   // ---------- 网络 17 ----------
   // 标题：请开始换夹具...
   // 含义：将 (#ChangeTool.S15 AND #StatusIn.do_ChgGrp_Pos) OR (#ChangeTool.S15 AND #ChangeTool.S17) 赋给 #ChangeTool.S17
   #ChangeTool.S17 := (#ChangeTool.S15 AND #StatusIn.do_ChgGrp_Pos) OR (#ChangeTool.S15 AND #ChangeTool.S17);
   // 含义：将 #ChangeTool.S15 AND NOT (#ChangeTool.S17) 赋给 "DB1146_PromptFree".Public.do_ChgGrp_Pos
   "DB1146_PromptFree".Public.do_ChgGrp_Pos := #ChangeTool.S15 AND NOT (#ChangeTool.S17);

   // ---------- 网络 18 ----------
   // 标题：快换盘锁紧 254放爪 253取爪
   // 含义：条件 ((#ChangeTool.S17 AND NOT (#ChangeTool.S19)) AND ("DB1080_Component".Robot.CTRL_IN.ProgNo = 253)) 成立时，将 TRUE 传送到 "DB1081_ValveCall".ST01.Z07.ExtAuto
   IF ((#ChangeTool.S17 AND NOT (#ChangeTool.S19)) AND ("DB1080_Component".Robot.CTRL_IN.ProgNo = 253)) THEN
       "DB1081_ValveCall".ST01.Z07.ExtAuto := TRUE;
   END_IF;
   // 含义：条件 ((#ChangeTool.S17 AND NOT (#ChangeTool.S19)) AND ("DB1080_Component".Robot.CTRL_IN.ProgNo = 254)) 成立时，将 TRUE 传送到 "DB1081_ValveCall".ST01.Z07.RetAuto
   IF ((#ChangeTool.S17 AND NOT (#ChangeTool.S19)) AND ("DB1080_Component".Robot.CTRL_IN.ProgNo = 254)) THEN
       "DB1081_ValveCall".ST01.Z07.RetAuto := TRUE;
   END_IF;
   // 含义：条件 #ChangeTool.S17 AND NOT (#ChangeTool.S19) 成立时，将 TRUE 传送到 "DB1060_AutoStep".Status.FirstStart
   IF #ChangeTool.S17 AND NOT (#ChangeTool.S19) THEN
       "DB1060_AutoStep".Status.FirstStart := TRUE;
   END_IF;
   // 含义：将 (((#ChangeTool.S17 AND ("DB1080_Component".Robot.CTRL_IN.ProgNo = 253))) AND "DB1081_ValveCall".ST01.Z07.ExtPos) OR (((#ChangeTool.S17 AND ("DB1080_Component".Robot.CTRL_IN.ProgNo = 254))) AND "DB1081_ValveCall".ST01.Z07.RetPos) OR (#ChangeTool.S17 AND #ChangeTool.S19) 赋给 #ChangeTool.S19
   #ChangeTool.S19 := (((#ChangeTool.S17 AND ("DB1080_Component".Robot.CTRL_IN.ProgNo = 253))) AND "DB1081_ValveCall".ST01.Z07.ExtPos) OR (((#ChangeTool.S17 AND ("DB1080_Component".Robot.CTRL_IN.ProgNo = 254))) AND "DB1081_ValveCall".ST01.Z07.RetPos) OR (#ChangeTool.S17 AND #ChangeTool.S19);

   // ---------- 网络 19 ----------
   // 标题：换爪完成确认
   // 含义：将 #ChangeTool.S19 AND NOT (#ChangeTool.S20) 赋给 #CmdOut.di_ChgGrp_Ack
   #CmdOut.di_ChgGrp_Ack := #ChangeTool.S19 AND NOT (#ChangeTool.S20);
   // 含义：将 #ChangeTool.S19 AND NOT (#ChangeTool.S20) 赋给 "DB1146_PromptFree".Public.do_ChgGrp_Act
   "DB1146_PromptFree".Public.do_ChgGrp_Act := #ChangeTool.S19 AND NOT (#ChangeTool.S20);
   // 含义：条件 (#ChangeTool.S19 AND NOT (#ChangeTool.S20)) AND NOT ("IToolAtPos") 成立时，将 TRUE 传送到 "DB1081_ValveCall".ST01.Z07.VentValveAuto
   IF (#ChangeTool.S19 AND NOT (#ChangeTool.S20)) AND NOT ("IToolAtPos") THEN
       "DB1081_ValveCall".ST01.Z07.VentValveAuto := TRUE;
   END_IF;
   // 含义：条件 #ChangeTool.S19 AND NOT (#ChangeTool.S20) 成立时，将 TRUE 传送到 "DB1081_ValveCall".ST01.Z08.RetAuto
   IF #ChangeTool.S19 AND NOT (#ChangeTool.S20) THEN
       "DB1081_ValveCall".ST01.Z08.RetAuto := TRUE;
   END_IF;
   // 含义：将 (#ChangeTool.S19 AND #StatusIn.do_ChgGrp_Don) OR (#ChangeTool.S19 AND #ChangeTool.S20) 赋给 #ChangeTool.S20
   #ChangeTool.S20 := (#ChangeTool.S19 AND #StatusIn.do_ChgGrp_Don) OR (#ChangeTool.S19 AND #ChangeTool.S20);

   // ---------- 网络 20 ----------
   // 标题：夹具库枪位置不正确！
   // 注释：M29.0常1临时屏蔽I6.0信号 20230911
   // 含义：将 (((((#ChangeTool.S20 AND ("DB1080_Component".Robot.CTRL_IN.ProgNo = 254))) AND (#CmdOut.gi_ToolPosNo = 1))) AND NOT (#Aux.AStation_ToolAtPosT.Q)) OR (((((#ChangeTool.S20 AND ("DB1080_Component".Robot.CTRL_IN.ProgNo = 254))) AND (#CmdOut.gi_ToolPosNo = 2))) AND NOT (#Aux.BStation_ToolAtPosT.Q)) 赋给 "DB1148_PromptBeeper".ST01.PutToolPosNotOk
   "DB1148_PromptBeeper".ST01.PutToolPosNotOk := (((((#ChangeTool.S20 AND ("DB1080_Component".Robot.CTRL_IN.ProgNo = 254))) AND (#CmdOut.gi_ToolPosNo = 1))) AND NOT (#Aux.AStation_ToolAtPosT.Q)) OR (((((#ChangeTool.S20 AND ("DB1080_Component".Robot.CTRL_IN.ProgNo = 254))) AND (#CmdOut.gi_ToolPosNo = 2))) AND NOT (#Aux.BStation_ToolAtPosT.Q));
   // 含义：将 (((((#ChangeTool.S20 AND ("DB1080_Component".Robot.CTRL_IN.ProgNo = 254))) AND (#CmdOut.gi_ToolPosNo = 1))) AND #Aux.AStation_ToolAtPosT.Q) OR (((((#ChangeTool.S20 AND ("DB1080_Component".Robot.CTRL_IN.ProgNo = 254))) AND (#CmdOut.gi_ToolPosNo = 2))) AND #Aux.BStation_ToolAtPosT.Q) OR ((((#ChangeTool.S20 AND ("DB1080_Component".Robot.CTRL_IN.ProgNo = 253))) AND "DB1081_ValveCall".ST01.Z07.ExtPos) AND "IToolAtPos") OR (#ChangeTool.S20 AND #ChangeTool.S22) 赋给 #ChangeTool.S22
   #ChangeTool.S22 := (((((#ChangeTool.S20 AND ("DB1080_Component".Robot.CTRL_IN.ProgNo = 254))) AND (#CmdOut.gi_ToolPosNo = 1))) AND #Aux.AStation_ToolAtPosT.Q) OR (((((#ChangeTool.S20 AND ("DB1080_Component".Robot.CTRL_IN.ProgNo = 254))) AND (#CmdOut.gi_ToolPosNo = 2))) AND #Aux.BStation_ToolAtPosT.Q) OR ((((#ChangeTool.S20 AND ("DB1080_Component".Robot.CTRL_IN.ProgNo = 253))) AND "DB1081_ValveCall".ST01.Z07.ExtPos) AND "IToolAtPos") OR (#ChangeTool.S20 AND #ChangeTool.S22);

   // ---------- 网络 21 ----------
   // 标题：防尘盖夹紧缸
   // 含义：条件 ((((#ChangeTool.S22 AND NOT (#ChangeTool.S23)) AND ("DB1080_Component".Robot.CTRL_IN.ProgNo <> 254))) OR ((#ChangeTool.S22 AND NOT (#ChangeTool.S23)) AND TRUE)) AND #Aux.AStation_ToolAtPosT.Q 成立时，将 TRUE 传送到 "DB1081_ValveCall".ST01.Z03.RetAuto
   IF ((((#ChangeTool.S22 AND NOT (#ChangeTool.S23)) AND ("DB1080_Component".Robot.CTRL_IN.ProgNo <> 254))) OR ((#ChangeTool.S22 AND NOT (#ChangeTool.S23)) AND TRUE)) AND #Aux.AStation_ToolAtPosT.Q THEN
       "DB1081_ValveCall".ST01.Z03.RetAuto := TRUE;
   END_IF;
   // 含义：条件 ((((#ChangeTool.S22 AND NOT (#ChangeTool.S23)) AND ("DB1080_Component".Robot.CTRL_IN.ProgNo <> 254))) OR ((#ChangeTool.S22 AND NOT (#ChangeTool.S23)) AND TRUE)) AND #Aux.BStation_ToolAtPosT.Q 成立时，将 TRUE 传送到 "DB1081_ValveCall".ST01.Z04.RetAuto
   IF ((((#ChangeTool.S22 AND NOT (#ChangeTool.S23)) AND ("DB1080_Component".Robot.CTRL_IN.ProgNo <> 254))) OR ((#ChangeTool.S22 AND NOT (#ChangeTool.S23)) AND TRUE)) AND #Aux.BStation_ToolAtPosT.Q THEN
       "DB1081_ValveCall".ST01.Z04.RetAuto := TRUE;
   END_IF;
   // 含义：将 (((#ChangeTool.S22 AND "DB1081_ValveCall".ST01.Z03.RetPos) OR (#ChangeTool.S22 AND NOT (#Aux.AStation_ToolAtPosT.Q))) AND "DB1081_ValveCall".ST01.Z04.RetPos) OR (((#ChangeTool.S22 AND "DB1081_ValveCall".ST01.Z03.RetPos) OR (#ChangeTool.S22 AND NOT (#Aux.AStation_ToolAtPosT.Q))) AND NOT (#Aux.BStation_ToolAtPosT.Q)) OR ((#ChangeTool.S22 AND ("DB1080_Component".Robot.CTRL_IN.ProgNo = 254))) OR (#ChangeTool.S22 AND #ChangeTool.S23) 赋给 #ChangeTool.S23
   #ChangeTool.S23 := (((#ChangeTool.S22 AND "DB1081_ValveCall".ST01.Z03.RetPos) OR (#ChangeTool.S22 AND NOT (#Aux.AStation_ToolAtPosT.Q))) AND "DB1081_ValveCall".ST01.Z04.RetPos) OR (((#ChangeTool.S22 AND "DB1081_ValveCall".ST01.Z03.RetPos) OR (#ChangeTool.S22 AND NOT (#Aux.AStation_ToolAtPosT.Q))) AND NOT (#Aux.BStation_ToolAtPosT.Q)) OR ((#ChangeTool.S22 AND ("DB1080_Component".Robot.CTRL_IN.ProgNo = 254))) OR (#ChangeTool.S22 AND #ChangeTool.S23);

   // ---------- 网络 22 ----------
   // 标题：TaskDone
   // 含义：条件 ((#ChangeTool.S23 OR #ChangeTool.ErrEnd OR #ChangeTool.ByPass) AND NOT (#ChangeTool.S25)) AND NOT (#ChangeTool.ErrEnd) 成立时，将 TRUE 传送到 #ChangeTool.TaskIO
   IF ((#ChangeTool.S23 OR #ChangeTool.ErrEnd OR #ChangeTool.ByPass) AND NOT (#ChangeTool.S25)) AND NOT (#ChangeTool.ErrEnd) THEN
       #ChangeTool.TaskIO := TRUE;
   END_IF;
   // 含义：条件 ((#ChangeTool.S23 OR #ChangeTool.ErrEnd OR #ChangeTool.ByPass) AND NOT (#ChangeTool.S25)) AND #ChangeTool.ErrEnd 成立时，将 TRUE 传送到 #ChangeTool.TaskNIO
   IF ((#ChangeTool.S23 OR #ChangeTool.ErrEnd OR #ChangeTool.ByPass) AND NOT (#ChangeTool.S25)) AND #ChangeTool.ErrEnd THEN
       #ChangeTool.TaskNIO := TRUE;
   END_IF;
   // 含义：将 #ChangeTool.S23 OR #ChangeTool.ErrEnd OR #ChangeTool.ByPass 赋给 #ChangeTool.S25
   #ChangeTool.S25 := #ChangeTool.S23 OR #ChangeTool.ErrEnd OR #ChangeTool.ByPass;

   // ---------- 网络 23 ----------
   // 标题：结束
   // 含义：将 (#ChangeTool.S25 OR #ChangeTool.ErrEnd) AND NOT (#ChangeTool.StartCmd) 赋给 #ChangeTool.StepEnd
   #ChangeTool.StepEnd := (#ChangeTool.S25 OR #ChangeTool.ErrEnd) AND NOT (#ChangeTool.StartCmd);
   // 含义：将 #ChangeTool.S25 OR #ChangeTool.ErrEnd 赋给 #ChangeTool.TaskDone
   #ChangeTool.TaskDone := #ChangeTool.S25 OR #ChangeTool.ErrEnd;

   // ---------- 网络 24 ----------
   // 含义：将 FALSE 赋给 #ChangeTool.StartCmd
   #ChangeTool.StartCmd := FALSE;

   // ---------- 网络 25 ----------
   // （空白网络）

   // ---------- 网络 26 ----------
   // 标题：本工位必须要做(可能条件暂时不满足)
   // 含义：将 (((((#Ctrl_Out.RobotAction = 0) AND #Aux.ToolAtPos) AND "ManMode_M") AND ("DB1900_Communication_PC".Recv.ChooseProgNo = 4))) OR (((((#Ctrl_Out.RobotAction = 0) AND #Aux.ToolAtPos) AND "ManMode_M") AND ("DB1900_Communication_PC".Recv.ChooseProgNo = 5))) OR (((#Ctrl_Out.RobotAction = 0) AND #Aux.ToolAtPos) AND "ASMMode_M") 赋给 #CheckBit.OKToStart
   #CheckBit.OKToStart := (((((#Ctrl_Out.RobotAction = 0) AND #Aux.ToolAtPos) AND "ManMode_M") AND ("DB1900_Communication_PC".Recv.ChooseProgNo = 4))) OR (((((#Ctrl_Out.RobotAction = 0) AND #Aux.ToolAtPos) AND "ManMode_M") AND ("DB1900_Communication_PC".Recv.ChooseProgNo = 5))) OR (((#Ctrl_Out.RobotAction = 0) AND #Aux.ToolAtPos) AND "ASMMode_M");
   // 含义：条件 "DB1900_Communication_PC".Recv.CheckAiguilleTPPB AND "ManMode_M" 成立时，将 TRUE 传送到 #CheckBit.StartCmd
   IF "DB1900_Communication_PC".Recv.CheckAiguilleTPPB AND "ManMode_M" THEN
       #CheckBit.StartCmd := TRUE;
   END_IF;

   // ---------- 网络 27 ----------
   // 标题：*********************************检查批头Start*************************************
   // 含义：将 (((((((#CheckBit.StartCmd AND #CheckBit.OKToStart) OR #CheckBit.StepStart) AND "AllMode_M") AND "DB1900_Communication_PC".Recv.Z05RetTPPB) AND ("DB1900_Communication_PC".Recv.Current_2 < 0.5))) AND NOT ("DB1040_HomePos".Status.Running)) AND NOT (#CheckBit.StepEnd) 赋给 #CheckBit.StepStart
   #CheckBit.StepStart := (((((((#CheckBit.StartCmd AND #CheckBit.OKToStart) OR #CheckBit.StepStart) AND "AllMode_M") AND "DB1900_Communication_PC".Recv.Z05RetTPPB) AND ("DB1900_Communication_PC".Recv.Current_2 < 0.5))) AND NOT ("DB1040_HomePos".Status.Running)) AND NOT (#CheckBit.StepEnd);
   // 含义：将 (((((((#CheckBit.StartCmd AND #CheckBit.OKToStart) OR #CheckBit.StepStart) AND "AllMode_M") AND "DB1900_Communication_PC".Recv.Z05RetTPPB) AND ("DB1900_Communication_PC".Recv.Current_2 < 0.5))) AND NOT ("DB1040_HomePos".Status.Running)) AND NOT (#CheckBit.StepEnd) 赋给 #CheckBit.Busy
   #CheckBit.Busy := (((((((#CheckBit.StartCmd AND #CheckBit.OKToStart) OR #CheckBit.StepStart) AND "AllMode_M") AND "DB1900_Communication_PC".Recv.Z05RetTPPB) AND ("DB1900_Communication_PC".Recv.Current_2 < 0.5))) AND NOT ("DB1040_HomePos".Status.Running)) AND NOT (#CheckBit.StepEnd);
   // 含义：将 (((((((#CheckBit.StartCmd AND #CheckBit.OKToStart) OR #CheckBit.StepStart) AND "AllMode_M") AND "DB1900_Communication_PC".Recv.Z05RetTPPB) AND ("DB1900_Communication_PC".Recv.Current_2 < 0.5))) AND NOT ("DB1040_HomePos".Status.Running)) AND NOT (#CheckBit.StepEnd) 赋给 "DB1900_Communication_PC".Send.RobotCheck
   "DB1900_Communication_PC".Send.RobotCheck := (((((((#CheckBit.StartCmd AND #CheckBit.OKToStart) OR #CheckBit.StepStart) AND "AllMode_M") AND "DB1900_Communication_PC".Recv.Z05RetTPPB) AND ("DB1900_Communication_PC".Recv.Current_2 < 0.5))) AND NOT ("DB1040_HomePos".Status.Running)) AND NOT (#CheckBit.StepEnd);
   // 含义：条件 NOT ((((((((#CheckBit.StartCmd AND #CheckBit.OKToStart) OR #CheckBit.StepStart) AND "AllMode_M") AND "DB1900_Communication_PC".Recv.Z05RetTPPB) AND ("DB1900_Communication_PC".Recv.Current_2 < 0.5))) AND NOT ("DB1040_HomePos".Status.Running)) AND NOT (#CheckBit.StepEnd)) 成立时，将 FALSE 传送到 #CheckBit.ErrEnd
   IF NOT ((((((((#CheckBit.StartCmd AND #CheckBit.OKToStart) OR #CheckBit.StepStart) AND "AllMode_M") AND "DB1900_Communication_PC".Recv.Z05RetTPPB) AND ("DB1900_Communication_PC".Recv.Current_2 < 0.5))) AND NOT ("DB1040_HomePos".Status.Running)) AND NOT (#CheckBit.StepEnd)) THEN
       #CheckBit.ErrEnd := FALSE;
   END_IF;
   // 含义：条件 NOT ((((((((#CheckBit.StartCmd AND #CheckBit.OKToStart) OR #CheckBit.StepStart) AND "AllMode_M") AND "DB1900_Communication_PC".Recv.Z05RetTPPB) AND ("DB1900_Communication_PC".Recv.Current_2 < 0.5))) AND NOT ("DB1040_HomePos".Status.Running)) AND NOT (#CheckBit.StepEnd)) 成立时，将 FALSE 传送到 "DB1148_PromptBeeper".Public.ScrLenFault
   IF NOT ((((((((#CheckBit.StartCmd AND #CheckBit.OKToStart) OR #CheckBit.StepStart) AND "AllMode_M") AND "DB1900_Communication_PC".Recv.Z05RetTPPB) AND ("DB1900_Communication_PC".Recv.Current_2 < 0.5))) AND NOT ("DB1040_HomePos".Status.Running)) AND NOT (#CheckBit.StepEnd)) THEN
       "DB1148_PromptBeeper".Public.ScrLenFault := FALSE;
   END_IF;
   // 含义：条件 NOT ((((((((#CheckBit.StartCmd AND #CheckBit.OKToStart) OR #CheckBit.StepStart) AND "AllMode_M") AND "DB1900_Communication_PC".Recv.Z05RetTPPB) AND ("DB1900_Communication_PC".Recv.Current_2 < 0.5))) AND NOT ("DB1040_HomePos".Status.Running)) AND NOT (#CheckBit.StepEnd)) 成立时，将 FALSE 传送到 #CmdOut.di_ChkScrew_Ack
   IF NOT ((((((((#CheckBit.StartCmd AND #CheckBit.OKToStart) OR #CheckBit.StepStart) AND "AllMode_M") AND "DB1900_Communication_PC".Recv.Z05RetTPPB) AND ("DB1900_Communication_PC".Recv.Current_2 < 0.5))) AND NOT ("DB1040_HomePos".Status.Running)) AND NOT (#CheckBit.StepEnd)) THEN
       #CmdOut.di_ChkScrew_Ack := FALSE;
   END_IF;

   // ---------- 网络 28 ----------
   // 标题：初始化
   // 含义：条件 (#CheckBit.StepStart AND NOT (#CheckBit.ErrEnd)) AND NOT (#CheckBit.S1) 成立时，将 FALSE 传送到 #CheckBit.TaskIO
   IF (#CheckBit.StepStart AND NOT (#CheckBit.ErrEnd)) AND NOT (#CheckBit.S1) THEN
       #CheckBit.TaskIO := FALSE;
   END_IF;
   // 含义：条件 (#CheckBit.StepStart AND NOT (#CheckBit.ErrEnd)) AND NOT (#CheckBit.S1) 成立时，将 FALSE 传送到 #CheckBit.TaskNIO
   IF (#CheckBit.StepStart AND NOT (#CheckBit.ErrEnd)) AND NOT (#CheckBit.S1) THEN
       #CheckBit.TaskNIO := FALSE;
   END_IF;
   // 含义：将 #CheckBit.StepStart AND NOT (#CheckBit.ErrEnd) 赋给 #CheckBit.S1
   #CheckBit.S1 := #CheckBit.StepStart AND NOT (#CheckBit.ErrEnd);

   // ---------- 网络 29 ----------
   // 标题：判断条件
   // 含义：当 #CheckBit.S1 为 TRUE 时置位 #CheckBit.S2，否则复位（触点→线圈）
   IF #CheckBit.S1 THEN
       #CheckBit.S2 := TRUE;
   ELSE
       #CheckBit.S2 := FALSE;
   END_IF;

   // ---------- 网络 30 ----------
   // 标题：电源夹具ID号错误，请检查夹具！
   // 含义：将 (#CheckBit.S2 AND #Aux.ToolAtPos) OR (#CheckBit.S2 AND #CheckBit.S5) 赋给 #CheckBit.S5
   #CheckBit.S5 := (#CheckBit.S2 AND #Aux.ToolAtPos) OR (#CheckBit.S2 AND #CheckBit.S5);

   // ---------- 网络 31 ----------
   // 标题：推力气缸
   // 含义：条件 #CheckBit.S5 AND NOT (#CheckBit.S7) 成立时，将 TRUE 传送到 "DB1081_ValveCall".ST01.Z01.ExtAuto
   IF #CheckBit.S5 AND NOT (#CheckBit.S7) THEN
       "DB1081_ValveCall".ST01.Z01.ExtAuto := TRUE;
   END_IF;
   // 含义：条件 #CheckBit.S5 AND NOT (#CheckBit.S7) 成立时，将 TRUE 传送到 "DB1081_ValveCall".ST01.Z02.VentValveAuto
   IF #CheckBit.S5 AND NOT (#CheckBit.S7) THEN
       "DB1081_ValveCall".ST01.Z02.VentValveAuto := TRUE;
   END_IF;
   // 含义：条件 #CheckBit.S5 AND NOT (#CheckBit.S7) 成立时，将 TRUE 传送到 "DB1081_ValveCall".ST01.Z05.RetAuto
   IF #CheckBit.S5 AND NOT (#CheckBit.S7) THEN
       "DB1081_ValveCall".ST01.Z05.RetAuto := TRUE;
   END_IF;
   // 含义：条件 #CheckBit.S5 AND NOT (#CheckBit.S7) 成立时，将 TRUE 传送到 "DB1081_ValveCall".ST01.Z06.RetAuto
   IF #CheckBit.S5 AND NOT (#CheckBit.S7) THEN
       "DB1081_ValveCall".ST01.Z06.RetAuto := TRUE;
   END_IF;
   // 含义：条件 (((#CheckBit.S5 AND NOT (#CheckBit.S7)) AND (#CmdOut.gi_ToolTypeNo = 13))) AND TRUE 成立时，将 FALSE 传送到 "QCamCoverExt"
   IF (((#CheckBit.S5 AND NOT (#CheckBit.S7)) AND (#CmdOut.gi_ToolTypeNo = 13))) AND TRUE THEN
       "QCamCoverExt" := FALSE;
   END_IF;
   // 含义：条件 (((#CheckBit.S5 AND NOT (#CheckBit.S7)) AND (#CmdOut.gi_ToolTypeNo = 13))) AND TRUE 成立时，将 TRUE 传送到 "QCamCoverRet"
   IF (((#CheckBit.S5 AND NOT (#CheckBit.S7)) AND (#CmdOut.gi_ToolTypeNo = 13))) AND TRUE THEN
       "QCamCoverRet" := TRUE;
   END_IF;
   // 含义：条件 #CheckBit.S5 AND NOT (#CheckBit.S7) 成立时，将 TRUE 传送到 "DB1081_ValveCall".ST01.Z08.ExtAuto
   IF #CheckBit.S5 AND NOT (#CheckBit.S7) THEN
       "DB1081_ValveCall".ST01.Z08.ExtAuto := TRUE;
   END_IF;
   // 含义：条件 #CheckBit.S5 AND NOT (#CheckBit.S7) 成立时，将 0.15 传送到 "DB1080_Component".Aux.Pressure
   IF #CheckBit.S5 AND NOT (#CheckBit.S7) THEN
       "DB1080_Component".Aux.Pressure := 0.15;
   END_IF;
   // 含义：将 ((((#CheckBit.S5 AND "DB1900_Communication_PC".Recv.ParaWriteDone) AND "DB1081_ValveCall".ST01.Z05.RetPos) AND "DB1081_ValveCall".ST01.Z06.RetPos) AND "IZ02ExtPos") OR (#CheckBit.S5 AND #CheckBit.S7) 赋给 #CheckBit.S7
   #CheckBit.S7 := ((((#CheckBit.S5 AND "DB1900_Communication_PC".Recv.ParaWriteDone) AND "DB1081_ValveCall".ST01.Z05.RetPos) AND "DB1081_ValveCall".ST01.Z06.RetPos) AND "IZ02ExtPos") OR (#CheckBit.S5 AND #CheckBit.S7);

   // ---------- 网络 32 ----------
   // 标题：数据写入 零点推力压缩量传递
   // 含义：条件 #CheckBit.S7 AND NOT (#CheckBit.S9) 成立时，将 "DB1900_Communication_PC".Para.ZeroPos 传送到 #Aux.ZeroPos
   IF #CheckBit.S7 AND NOT (#CheckBit.S9) THEN
       #Aux.ZeroPos := "DB1900_Communication_PC".Para.ZeroPos;
   END_IF;
   // 含义：当 #CheckBit.S7 为 TRUE 时置位 #CheckBit.S9，否则复位（触点→线圈）
   IF #CheckBit.S7 THEN
       #CheckBit.S9 := TRUE;
   ELSE
       #CheckBit.S9 := FALSE;
   END_IF;

   // ---------- 网络 33 ----------
   // 含义：将 (#CheckBit.S9 AND NOT ("DB1080_Component".Robot.Status.Busy)) OR (#CheckBit.S9 AND #CheckBit.S10) 赋给 #CheckBit.S10
   #CheckBit.S10 := (#CheckBit.S9 AND NOT ("DB1080_Component".Robot.Status.Busy)) OR (#CheckBit.S9 AND #CheckBit.S10);

   // ---------- 网络 34 ----------
   // 标题：调用机器人
   // 含义：条件 (#CheckBit.S10 OR #CheckBit.S9) AND NOT (#CheckBit.S15) 成立时，将 TRUE 传送到 "DB1080_Component".Robot.Cmd.Auto.ProgStart
   IF (#CheckBit.S10 OR #CheckBit.S9) AND NOT (#CheckBit.S15) THEN
       "DB1080_Component".Robot.Cmd.Auto.ProgStart := TRUE;
   END_IF;
   // 含义：条件 (#CheckBit.S10 OR #CheckBit.S9) AND NOT (#CheckBit.S15) 成立时，将 40 传送到 "DB1080_Component".Robot.CTRL_IN.RobotSpeed
   IF (#CheckBit.S10 OR #CheckBit.S9) AND NOT (#CheckBit.S15) THEN
       "DB1080_Component".Robot.CTRL_IN.RobotSpeed := 40;
   END_IF;
   // 含义：条件 ((#CheckBit.S10 OR #CheckBit.S9) AND NOT (#CheckBit.S15)) AND "ASMMode_M" 成立时，将 4 传送到 "DB1080_Component".Robot.CTRL_IN.ProgNo
   IF ((#CheckBit.S10 OR #CheckBit.S9) AND NOT (#CheckBit.S15)) AND "ASMMode_M" THEN
       "DB1080_Component".Robot.CTRL_IN.ProgNo := 4;
   END_IF;
   // 含义：条件 ((((((#CheckBit.S10 OR #CheckBit.S9) AND NOT (#CheckBit.S15)) AND "ManMode_M") AND ("DB1900_Communication_PC".Recv.ChooseProgNo = 5))) AND (#Aux.CheckNo = 1)) 成立时，将 TRUE 传送到 "DB1081_ValveCall".ST01.Z02.RetAuto
   IF ((((((#CheckBit.S10 OR #CheckBit.S9) AND NOT (#CheckBit.S15)) AND "ManMode_M") AND ("DB1900_Communication_PC".Recv.ChooseProgNo = 5))) AND (#Aux.CheckNo = 1)) THEN
       "DB1081_ValveCall".ST01.Z02.RetAuto := TRUE;
   END_IF;
   // 含义：条件 ((((((#CheckBit.S10 OR #CheckBit.S9) AND NOT (#CheckBit.S15)) AND "ManMode_M") AND ("DB1900_Communication_PC".Recv.ChooseProgNo = 5))) AND (#Aux.CheckNo = 1)) 成立时，将 10 传送到 "DB1080_Component".Robot.CTRL_IN.ProgNo
   IF ((((((#CheckBit.S10 OR #CheckBit.S9) AND NOT (#CheckBit.S15)) AND "ManMode_M") AND ("DB1900_Communication_PC".Recv.ChooseProgNo = 5))) AND (#Aux.CheckNo = 1)) THEN
       "DB1080_Component".Robot.CTRL_IN.ProgNo := 10;
   END_IF;
   // 含义：条件 ((((((#CheckBit.S10 OR #CheckBit.S9) AND NOT (#CheckBit.S15)) AND "ManMode_M") AND ("DB1900_Communication_PC".Recv.ChooseProgNo = 5))) AND (#Aux.CheckNo = 2)) 成立时，将 TRUE 传送到 "DB1081_ValveCall".ST01.Z02.VentValveAuto
   IF ((((((#CheckBit.S10 OR #CheckBit.S9) AND NOT (#CheckBit.S15)) AND "ManMode_M") AND ("DB1900_Communication_PC".Recv.ChooseProgNo = 5))) AND (#Aux.CheckNo = 2)) THEN
       "DB1081_ValveCall".ST01.Z02.VentValveAuto := TRUE;
   END_IF;
   // 含义：条件 ((((((#CheckBit.S10 OR #CheckBit.S9) AND NOT (#CheckBit.S15)) AND "ManMode_M") AND ("DB1900_Communication_PC".Recv.ChooseProgNo = 5))) AND (#Aux.CheckNo = 2)) 成立时，将 11 传送到 "DB1080_Component".Robot.CTRL_IN.ProgNo
   IF ((((((#CheckBit.S10 OR #CheckBit.S9) AND NOT (#CheckBit.S15)) AND "ManMode_M") AND ("DB1900_Communication_PC".Recv.ChooseProgNo = 5))) AND (#Aux.CheckNo = 2)) THEN
       "DB1080_Component".Robot.CTRL_IN.ProgNo := 11;
   END_IF;
   // 含义：条件 ((((((#CheckBit.S10 OR #CheckBit.S9) AND NOT (#CheckBit.S15)) AND "ManMode_M") AND ("DB1900_Communication_PC".Recv.ChooseProgNo = 5))) AND (#Aux.CheckNo = 3)) 成立时，将 TRUE 传送到 "DB1081_ValveCall".ST01.Z01.ExtAuto
   IF ((((((#CheckBit.S10 OR #CheckBit.S9) AND NOT (#CheckBit.S15)) AND "ManMode_M") AND ("DB1900_Communication_PC".Recv.ChooseProgNo = 5))) AND (#Aux.CheckNo = 3)) THEN
       "DB1081_ValveCall".ST01.Z01.ExtAuto := TRUE;
   END_IF;
   // 含义：条件 ((((((#CheckBit.S10 OR #CheckBit.S9) AND NOT (#CheckBit.S15)) AND "ManMode_M") AND ("DB1900_Communication_PC".Recv.ChooseProgNo = 5))) AND (#Aux.CheckNo = 3)) 成立时，将 TRUE 传送到 "DB1081_ValveCall".ST01.Z02.RetAuto
   IF ((((((#CheckBit.S10 OR #CheckBit.S9) AND NOT (#CheckBit.S15)) AND "ManMode_M") AND ("DB1900_Communication_PC".Recv.ChooseProgNo = 5))) AND (#Aux.CheckNo = 3)) THEN
       "DB1081_ValveCall".ST01.Z02.RetAuto := TRUE;
   END_IF;
   // 含义：条件 ((((((#CheckBit.S10 OR #CheckBit.S9) AND NOT (#CheckBit.S15)) AND "ManMode_M") AND ("DB1900_Communication_PC".Recv.ChooseProgNo = 5))) AND (#Aux.CheckNo = 3)) 成立时，将 12 传送到 "DB1080_Component".Robot.CTRL_IN.ProgNo
   IF ((((((#CheckBit.S10 OR #CheckBit.S9) AND NOT (#CheckBit.S15)) AND "ManMode_M") AND ("DB1900_Communication_PC".Recv.ChooseProgNo = 5))) AND (#Aux.CheckNo = 3)) THEN
       "DB1080_Component".Robot.CTRL_IN.ProgNo := 12;
   END_IF;
   // 含义：将 ((#CheckBit.S10 OR #CheckBit.S9) AND "DB1080_Component".Robot.Status.Busy) OR ((#CheckBit.S10 OR #CheckBit.S9) AND #CheckBit.S15) 赋给 #CheckBit.S15
   #CheckBit.S15 := ((#CheckBit.S10 OR #CheckBit.S9) AND "DB1080_Component".Robot.Status.Busy) OR ((#CheckBit.S10 OR #CheckBit.S9) AND #CheckBit.S15);

   // ---------- 网络 35 ----------
   // 含义：将 (#CheckBit.S15 AND #StatusIn.do_ChkScrew_Act) OR (#CheckBit.S15 AND #CheckBit.S17) 赋给 #CheckBit.S17
   #CheckBit.S17 := (#CheckBit.S15 AND #StatusIn.do_ChkScrew_Act) OR (#CheckBit.S15 AND #CheckBit.S17);
   // 含义：将 #CheckBit.S15 AND NOT (#CheckBit.S17) 赋给 "DB1146_PromptFree".Public.do_ChkScrew_Act
   "DB1146_PromptFree".Public.do_ChkScrew_Act := #CheckBit.S15 AND NOT (#CheckBit.S17);

   // ---------- 网络 36 ----------
   // 标题：初始化
   // 含义：条件 (#CheckBit.S17 AND NOT (#CheckBit.S19)) AND #StatusIn.do_ChkScrew_Pos 成立时，将 (#Aux.ZeroPos - #Aux.go_X) 传送到 #Aux.ScrLen
   IF (#CheckBit.S17 AND NOT (#CheckBit.S19)) AND #StatusIn.do_ChkScrew_Pos THEN
       #Aux.ScrLen := (#Aux.ZeroPos - #Aux.go_X);
   END_IF;
   // 含义：将 (#CheckBit.S17 AND NOT (#CheckBit.S19)) AND #StatusIn.do_ChkScrew_Pos 赋给 "DB1146_PromptFree".Public.AskPcData_1
   "DB1146_PromptFree".Public.AskPcData_1 := (#CheckBit.S17 AND NOT (#CheckBit.S19)) AND #StatusIn.do_ChkScrew_Pos;
   // 含义：条件 ((#CheckBit.S17 AND NOT (#CheckBit.S19)) AND ("DB1080_Component".ClinyderPos.Ctrl_Out.Cur_Val_Out > 0.5)) 成立时，将 20 传送到 "DB1080_Component".Robot.CTRL_IN.RobotSpeed
   IF ((#CheckBit.S17 AND NOT (#CheckBit.S19)) AND ("DB1080_Component".ClinyderPos.Ctrl_Out.Cur_Val_Out > 0.5)) THEN
       "DB1080_Component".Robot.CTRL_IN.RobotSpeed := 20;
   END_IF;
   // 含义：条件 ((#CheckBit.S17 AND NOT (#CheckBit.S19)) AND ("DB1080_Component".ClinyderPos.Ctrl_Out.Cur_Val_Out < 0.5)) 成立时，将 50 传送到 "DB1080_Component".Robot.CTRL_IN.RobotSpeed
   IF ((#CheckBit.S17 AND NOT (#CheckBit.S19)) AND ("DB1080_Component".ClinyderPos.Ctrl_Out.Cur_Val_Out < 0.5)) THEN
       "DB1080_Component".Robot.CTRL_IN.RobotSpeed := 50;
   END_IF;
   // 含义：将 (#CheckBit.S17 AND "DB1900_Communication_PC".Recv.ParaWriteDone) OR (#CheckBit.S17 AND #CheckBit.S23) 赋给 #CheckBit.S23
   #CheckBit.S23 := (#CheckBit.S17 AND "DB1900_Communication_PC".Recv.ParaWriteDone) OR (#CheckBit.S17 AND #CheckBit.S23);

   // ---------- 网络 37 ----------
   // 标题：**********************计算************************
   // 含义：本网络为 StructuredText（SCL）原文重建，非 LAD 折叠
   IF #CheckBit.S23 AND #StatusIn.do_ChkScrew_Pos AND
       ("DB1900_Communication_PC".Recv.ChooseProgNo = 4 OR "AutoMode_M") AND
       NOT #CheckBit.S25
   THEN
       IF #Aux.ZeroPos - #Aux.go_X > "DB1900_Communication_PC".Para.ScrLen - 15 AND
           #Aux.ZeroPos - #Aux.go_X < "DB1900_Communication_PC".Para.ScrLen + 15
       THEN
           "DB1148_PromptBeeper".Public.ScrLenFault := false;
           #CmdOut.di_ChkScrew_Ack := true;
       ELSE
           "DB1148_PromptBeeper".Public.ScrLenFault := true;
       END_IF;
   END_IF;
   "R_TRIG_DB"(CLK := #CmdOut.di_Front_Sig AND #CheckBit.S23 AND #StatusIn.do_ChkScrew_Pos,
               Q => #EdgeDetc.Pulse[0]);
   IF #EdgeDetc.Pulse[0]
   THEN
       "DB1900_Communication_PC".Send.ScrTestLen := #Aux.ZeroPos - #Aux.go_X;
   END_IF;

   // ---------- 网络 38 ----------
   // 标题：完成确认
   // 含义：将 (#CheckBit.S23 AND #StatusIn.do_ChkScrew_Don) OR (#CheckBit.S23 AND #CheckBit.S25) 赋给 #CheckBit.S25
   #CheckBit.S25 := (#CheckBit.S23 AND #StatusIn.do_ChkScrew_Don) OR (#CheckBit.S23 AND #CheckBit.S25);
   // 含义：条件 #CheckBit.S23 AND #CmdOut.di_ChkScrew_Ack 成立时，将 FALSE 传送到 "DB1148_PromptBeeper".Public.ScrLenFault
   IF #CheckBit.S23 AND #CmdOut.di_ChkScrew_Ack THEN
       "DB1148_PromptBeeper".Public.ScrLenFault := FALSE;
   END_IF;
   // 含义：条件 ((#CheckBit.S23 AND NOT (#CheckBit.S25)) AND ("DB1900_Communication_PC".Recv.ChooseProgNo = 5)) 成立时，将 TRUE 传送到 #CmdOut.di_ChkScrew_Ack
   IF ((#CheckBit.S23 AND NOT (#CheckBit.S25)) AND ("DB1900_Communication_PC".Recv.ChooseProgNo = 5)) THEN
       #CmdOut.di_ChkScrew_Ack := TRUE;
   END_IF;
   // 含义：条件 ((#CheckBit.S23 AND NOT (#CheckBit.S25)) AND "DB1148_PromptBeeper".Public.ScrLenFault) AND "ErrRst_M" 成立时，将 TRUE 传送到 #CheckBit.ErrEnd
   IF ((#CheckBit.S23 AND NOT (#CheckBit.S25)) AND "DB1148_PromptBeeper".Public.ScrLenFault) AND "ErrRst_M" THEN
       #CheckBit.ErrEnd := TRUE;
   END_IF;

   // ---------- 网络 39 ----------
   // 标题：推力气缸
   // 含义：条件 #CheckBit.S25 AND NOT (#CheckBit.S27) 成立时，将 TRUE 传送到 "DB1081_ValveCall".ST01.Z01.ExtAuto
   IF #CheckBit.S25 AND NOT (#CheckBit.S27) THEN
       "DB1081_ValveCall".ST01.Z01.ExtAuto := TRUE;
   END_IF;
   // 含义：条件 #CheckBit.S25 AND NOT (#CheckBit.S27) 成立时，将 TRUE 传送到 "DB1081_ValveCall".ST01.Z02.VentValveAuto
   IF #CheckBit.S25 AND NOT (#CheckBit.S27) THEN
       "DB1081_ValveCall".ST01.Z02.VentValveAuto := TRUE;
   END_IF;
   // 含义：条件 #CheckBit.S25 AND NOT (#CheckBit.S27) 成立时，将 0.3 传送到 "DB1080_Component".Aux.Pressure
   IF #CheckBit.S25 AND NOT (#CheckBit.S27) THEN
       "DB1080_Component".Aux.Pressure := 0.3;
   END_IF;
   // 含义：条件 #CheckBit.S25 AND NOT (#CheckBit.S27) 成立时，将 TRUE 传送到 "DB1081_ValveCall".ST01.Z08.RetAuto
   IF #CheckBit.S25 AND NOT (#CheckBit.S27) THEN
       "DB1081_ValveCall".ST01.Z08.RetAuto := TRUE;
   END_IF;
   // 含义：将 ((#CheckBit.S25 AND "DB1081_ValveCall".ST01.Z01.ExtPos) AND "DB1081_ValveCall".ST01.Z02.VentValve) OR (#CheckBit.S25 AND #CheckBit.S27) 赋给 #CheckBit.S27
   #CheckBit.S27 := ((#CheckBit.S25 AND "DB1081_ValveCall".ST01.Z01.ExtPos) AND "DB1081_ValveCall".ST01.Z02.VentValve) OR (#CheckBit.S25 AND #CheckBit.S27);

   // ---------- 网络 40 ----------
   // 标题：TaskDone
   // 含义：条件 ((#CheckBit.S27 OR #CheckBit.ErrEnd OR #CheckBit.ByPass) AND NOT (#CheckBit.S32)) AND NOT (#CheckBit.ErrEnd) 成立时，将 TRUE 传送到 #CheckBit.TaskIO
   IF ((#CheckBit.S27 OR #CheckBit.ErrEnd OR #CheckBit.ByPass) AND NOT (#CheckBit.S32)) AND NOT (#CheckBit.ErrEnd) THEN
       #CheckBit.TaskIO := TRUE;
   END_IF;
   // 含义：条件 ((#CheckBit.S27 OR #CheckBit.ErrEnd OR #CheckBit.ByPass) AND NOT (#CheckBit.S32)) AND #CheckBit.ErrEnd 成立时，将 TRUE 传送到 #CheckBit.TaskNIO
   IF ((#CheckBit.S27 OR #CheckBit.ErrEnd OR #CheckBit.ByPass) AND NOT (#CheckBit.S32)) AND #CheckBit.ErrEnd THEN
       #CheckBit.TaskNIO := TRUE;
   END_IF;
   // 含义：条件 (#CheckBit.S27 OR #CheckBit.ErrEnd OR #CheckBit.ByPass) AND NOT (#CheckBit.S32) 成立时，将 TRUE 传送到 "DB1081_ValveCall".ST01.Z08.RetAuto
   IF (#CheckBit.S27 OR #CheckBit.ErrEnd OR #CheckBit.ByPass) AND NOT (#CheckBit.S32) THEN
       "DB1081_ValveCall".ST01.Z08.RetAuto := TRUE;
   END_IF;
   // 含义：条件 (#CheckBit.S27 OR #CheckBit.ErrEnd OR #CheckBit.ByPass) AND NOT (#CheckBit.S32) 成立时，将 FALSE 传送到 "DB1060_AutoStep".Status.FirstStart
   IF (#CheckBit.S27 OR #CheckBit.ErrEnd OR #CheckBit.ByPass) AND NOT (#CheckBit.S32) THEN
       "DB1060_AutoStep".Status.FirstStart := FALSE;
   END_IF;
   // 含义：条件 (#CheckBit.S27 OR #CheckBit.ErrEnd OR #CheckBit.ByPass) AND NOT (#CheckBit.S32) 成立时，将 20 传送到 "DB1080_Component".Robot.CTRL_IN.RobotSpeed
   IF (#CheckBit.S27 OR #CheckBit.ErrEnd OR #CheckBit.ByPass) AND NOT (#CheckBit.S32) THEN
       "DB1080_Component".Robot.CTRL_IN.RobotSpeed := 20;
   END_IF;
   // 含义：将 #CheckBit.S27 OR #CheckBit.ErrEnd OR #CheckBit.ByPass 赋给 #CheckBit.S32
   #CheckBit.S32 := #CheckBit.S27 OR #CheckBit.ErrEnd OR #CheckBit.ByPass;

   // ---------- 网络 41 ----------
   // 标题：结束
   // 含义：将 (#CheckBit.S32 OR #CheckBit.ErrEnd) AND NOT (#CheckBit.StartCmd) 赋给 #CheckBit.StepEnd
   #CheckBit.StepEnd := (#CheckBit.S32 OR #CheckBit.ErrEnd) AND NOT (#CheckBit.StartCmd);
   // 含义：将 #CheckBit.S32 OR #CheckBit.ErrEnd 赋给 #CheckBit.TaskDone
   #CheckBit.TaskDone := #CheckBit.S32 OR #CheckBit.ErrEnd;

   // ---------- 网络 42 ----------
   // 含义：将 FALSE 赋给 #CheckBit.StartCmd
   #CheckBit.StartCmd := FALSE;
END_FUNCTION_BLOCK

FUNCTION_BLOCK "FB1060_AutoStep"   // FB1060, SCL
{ S7_Optimized_Access := 'FALSE' }
// ============================================================
//  Block: FB1060_AutoStep
//  ============================================================
//  编号：FB1060
//  原始语言：LAD（规则翻译为 SCL）
//  含义：自动循环起点
   VAR
      Status : Struct   // 状态
         Running : Bool;   // 自动运行中
         OkToStart : Bool;   // 设备可以启动
         FirstStart : Bool;   // 换枪后第一次
      END_STRUCT;
      Aux : Struct   // 静态变量
         HoleNo : Int;   // 工作流程数
      END_STRUCT;
      EdgeDetc : Struct   // 静态变量
         Pulse : Array[0..15] of Bool;   // 静态变量
      END_STRUCT;
      MainStep : "UDT_Step";   // 自动流程步
      CycleTime : "FB5008_CycleTime";   // 静态变量
      RobotAutoStep : "FB1061_RobotAutoStep";   // 静态变量
      HorDrillAutoStep : "FB1062_HorDrillAutoStep";   // 静态变量
      DownDrillAutoStep : "FB1063_DownDrillAutoStep";   // 静态变量
      DiamondAutoStep : "FB1064_DiamondAutostep";   // 静态变量
   END_VAR
   VAR_TEMP
      StepPls : Bool;
   END_VAR
BEGIN

   // ---------- 网络 1 ----------
   // 标题：模式分配
   // 含义：将 ("StepMode_M" AND "DB1001_SysMode".SubSysMode.Mode.StepPls) OR ("StepMode_M" AND #MainStep.StartCmd_ManMode) OR "ManMode_M" OR "AutoMode_M" 赋给 #StepPls
   #StepPls := ("StepMode_M" AND "DB1001_SysMode".SubSysMode.Mode.StepPls) OR ("StepMode_M" AND #MainStep.StartCmd_ManMode) OR "ManMode_M" OR "AutoMode_M";
   // 含义：条件 NOT ("AllMode_M") 成立时，将 TRUE 传送到 "DB1081_ValveCall".ST01.Z08.RetAuto
   IF NOT ("AllMode_M") THEN
       "DB1081_ValveCall".ST01.Z08.RetAuto := TRUE;
   END_IF;
   // 含义：当 "DB1900_Communication_PC".Recv.EmmMode 为 TRUE 时置位 "DB1148_PromptBeeper".Public.PcErr，否则复位（触点→线圈）
   IF "DB1900_Communication_PC".Recv.EmmMode THEN
       "DB1148_PromptBeeper".Public.PcErr := TRUE;
   ELSE
       "DB1148_PromptBeeper".Public.PcErr := FALSE;
   END_IF;
   // 含义：调用计数器实例 "Timer_RecvEmmMode".TON（上升沿计数，当前值写入 CV）
   "Timer_RecvEmmMode".TON(IN := "DB1900_Communication_PC".Recv.EmmMode,
                           PT := T#5s);
   // 含义：条件 "Timer_RecvEmmMode".Q 成立时，将 TRUE 传送到 "DB1900_Communication_PC".Send.PowerOff
   IF "Timer_RecvEmmMode".Q THEN
       "DB1900_Communication_PC".Send.PowerOff := TRUE;
   END_IF;
   // 含义：条件 "DB1900_Communication_PC".Recv.EmmMode 成立时，将 TRUE 传送到 "DB1080_Component".Robot.Cmd.Auto.Stop
   IF "DB1900_Communication_PC".Recv.EmmMode THEN
       "DB1080_Component".Robot.Cmd.Auto.Stop := TRUE;
   END_IF;
   // 含义：条件 "DB1900_Communication_PC".Recv.EmmMode 成立时，将 0 传送到 "DB1080_Component".Robot.CTRL_IN.ProgNo
   IF "DB1900_Communication_PC".Recv.EmmMode THEN
       "DB1080_Component".Robot.CTRL_IN.ProgNo := 0;
   END_IF;
   // 含义：条件 "DB1900_Communication_PC".Recv.PosNoClear OR "DB1900_Communication_PC".Recv.ClearHoleNoReq OR (("DB720_KuKa_MainCtrl".CmdOut.gi_ToolTypeNo = 2) AND "DB1900_Communication_PC".Recv.ChangeTool) 成立时，将 0 传送到 #Aux.HoleNo
   IF "DB1900_Communication_PC".Recv.PosNoClear OR "DB1900_Communication_PC".Recv.ClearHoleNoReq OR (("DB720_KuKa_MainCtrl".CmdOut.gi_ToolTypeNo = 2) AND "DB1900_Communication_PC".Recv.ChangeTool) THEN
       #Aux.HoleNo := 0;
   END_IF;
   // 含义：将 #Aux.HoleNo 赋给 "DB1900_Communication_PC".Send.PosNo
   "DB1900_Communication_PC".Send.PosNo := #Aux.HoleNo;
   // 含义：将 #Aux.HoleNo 赋给 "DB1900_Communication_PC".Send.HoleNo
   "DB1900_Communication_PC".Send.HoleNo := #Aux.HoleNo;
   // 含义：将 ("DB1900_Communication_PC".Recv.ClearHoleNoReq AND (#Aux.HoleNo = 0)) 赋给 "DB1900_Communication_PC".Send.ClearHoleNum
   "DB1900_Communication_PC".Send.ClearHoleNum := ("DB1900_Communication_PC".Recv.ClearHoleNoReq AND (#Aux.HoleNo = 0));
   // 含义：将 (("DB1900_Communication_PC".Para.DrillDirection1 OR "DB1900_Communication_PC".Para.DrillDirection3) AND ("DB1900_Communication_PC".Para.Auto_Force[5] = 0.0)) 赋给 "DB1148_PromptBeeper".Public.ForceCannotZero
   "DB1148_PromptBeeper".Public.ForceCannotZero := (("DB1900_Communication_PC".Para.DrillDirection1 OR "DB1900_Communication_PC".Para.DrillDirection3) AND ("DB1900_Communication_PC".Para.Auto_Force[5] = 0.0));
   // 含义：条件 "ManMode_M" AND "ErrRst_M" 成立时，将 FALSE 传送到 "DB1900_Communication_PC".Send.PowerOff
   IF "ManMode_M" AND "ErrRst_M" THEN
       "DB1900_Communication_PC".Send.PowerOff := FALSE;
   END_IF;
   // 含义：条件 "ManMode_M" AND "ErrRst_M" 成立时，将 FALSE 传送到 "DB1147_PromptStartNotPmt".Public.ParaWiriteOuttime
   IF "ManMode_M" AND "ErrRst_M" THEN
       "DB1147_PromptStartNotPmt".Public.ParaWiriteOuttime := FALSE;
   END_IF;
   // 含义：条件 "ManMode_M" AND "ErrRst_M" 成立时，将 FALSE 传送到 "DB1148_PromptBeeper".Public.BitStuckErr_Fixture
   IF "ManMode_M" AND "ErrRst_M" THEN
       "DB1148_PromptBeeper".Public.BitStuckErr_Fixture := FALSE;
   END_IF;
   // 含义：条件 "ManMode_M" AND "ErrRst_M" 成立时，将 FALSE 传送到 "DB1148_PromptBeeper".Public.BitStuckErr_HighCurrent
   IF "ManMode_M" AND "ErrRst_M" THEN
       "DB1148_PromptBeeper".Public.BitStuckErr_HighCurrent := FALSE;
   END_IF;
   // 含义：条件 "ManMode_M" AND "ErrRst_M" 成立时，将 FALSE 传送到 "DB1148_PromptBeeper".Public.DiamondCoreNOK
   IF "ManMode_M" AND "ErrRst_M" THEN
       "DB1148_PromptBeeper".Public.DiamondCoreNOK := FALSE;
   END_IF;
   // 含义：条件 "ManMode_M" AND "ErrRst_M" 成立时，将 FALSE 传送到 "DB1147_PromptStartNotPmt".Public.PcCommErr
   IF "ManMode_M" AND "ErrRst_M" THEN
       "DB1147_PromptStartNotPmt".Public.PcCommErr := FALSE;
   END_IF;

   // ---------- 网络 2 ----------
   // 标题：Running;
   // 含义：将 ((((NOT ("DB1001_SysMode".SubSysMode.Status.ErrPresent) AND "DB1040_HomePos".Status.AllStationInHomePos) AND "AutoMode_M") AND "IAutoModeStart") OR #Status.Running) AND "ASMMode_M" 赋给 #Status.Running
   #Status.Running := ((((NOT ("DB1001_SysMode".SubSysMode.Status.ErrPresent) AND "DB1040_HomePos".Status.AllStationInHomePos) AND "AutoMode_M") AND "IAutoModeStart") OR #Status.Running) AND "ASMMode_M";

   // ---------- 网络 3 ----------
   // 标题：提示回原点
   // 含义：将 (("ASMMode_M" AND NOT (#Status.Running)) AND NOT ("DB1040_HomePos".Status.AllStationInHomePos)) AND NOT ("DB1040_HomePos".MainStep.Start) 赋给 "DB1147_PromptStartNotPmt".Public.ToBeHomePos
   "DB1147_PromptStartNotPmt".Public.ToBeHomePos := (("ASMMode_M" AND NOT (#Status.Running)) AND NOT ("DB1040_HomePos".Status.AllStationInHomePos)) AND NOT ("DB1040_HomePos".MainStep.Start);
   // 含义：将 "ASMMode_M" AND NOT ("DB1001_SysMode".SubSysMode.Status.ErrPresent) 赋给 #Status.OkToStart
   #Status.OkToStart := "ASMMode_M" AND NOT ("DB1001_SysMode".SubSysMode.Status.ErrPresent);

   // ---------- 网络 4 ----------
   // 标题：自动步开始
   // 注释：自动循环起点
   // 含义：将 (((((((#Status.OkToStart AND "IAutoModeStart") OR #MainStep.Start) AND #Status.Running) AND NOT ("DB1147_PromptStartNotPmt".Public.PcCommErr)) AND NOT ("DB1900_Communication_PC".Recv.EmmMode)) AND NOT ("DB1040_HomePos".MainStep.Start)) AND NOT (#MainStep.End)) AND NOT ("DB1900_Communication_PC".Send.PowerOff) 赋给 #MainStep.Start
   #MainStep.Start := (((((((#Status.OkToStart AND "IAutoModeStart") OR #MainStep.Start) AND #Status.Running) AND NOT ("DB1147_PromptStartNotPmt".Public.PcCommErr)) AND NOT ("DB1900_Communication_PC".Recv.EmmMode)) AND NOT ("DB1040_HomePos".MainStep.Start)) AND NOT (#MainStep.End)) AND NOT ("DB1900_Communication_PC".Send.PowerOff);
   // 含义：条件 NOT ((#Status.OkToStart AND "IAutoModeStart") OR #MainStep.Start) 成立时，将 FALSE 传送到 #MainStep.ErrEnd
   IF NOT ((#Status.OkToStart AND "IAutoModeStart") OR #MainStep.Start) THEN
       #MainStep.ErrEnd := FALSE;
   END_IF;
   // 含义：条件 NOT ((#Status.OkToStart AND "IAutoModeStart") OR #MainStep.Start) 成立时，将 FALSE 传送到 "DB1900_Communication_PC".Send.DrillRunning
   IF NOT ((#Status.OkToStart AND "IAutoModeStart") OR #MainStep.Start) THEN
       "DB1900_Communication_PC".Send.DrillRunning := FALSE;
   END_IF;
   // 含义：条件 NOT ((#Status.OkToStart AND "IAutoModeStart") OR #MainStep.Start) 成立时，将 FALSE 传送到 #DiamondAutoStep.DiamondStep.StartCmd
   IF NOT ((#Status.OkToStart AND "IAutoModeStart") OR #MainStep.Start) THEN
       #DiamondAutoStep.DiamondStep.StartCmd := FALSE;
   END_IF;
   // 含义：调用定时器实例 "DB1042_Timer".FirstStartTime.TON
   "DB1042_Timer".FirstStartTime.TON(IN := NOT ((#Status.OkToStart AND "IAutoModeStart") OR #MainStep.Start),
                                     PT := T#6s);
   // 含义：条件 (NOT ((#Status.OkToStart AND "IAutoModeStart") OR #MainStep.Start)) AND "DB1042_Timer".FirstStartTime.Q 成立时，将 TRUE 传送到 #Status.FirstStart
   IF (NOT ((#Status.OkToStart AND "IAutoModeStart") OR #MainStep.Start)) AND "DB1042_Timer".FirstStartTime.Q THEN
       #Status.FirstStart := TRUE;
   END_IF;

   // ---------- 网络 5 ----------
   // 标题：有故障，断开正常流程，转入故障处理；
   // 含义：将 #MainStep.Start AND NOT (#MainStep.ErrEnd) 赋给 #MainStep.S1
   #MainStep.S1 := #MainStep.Start AND NOT (#MainStep.ErrEnd);

   // ---------- 网络 6 ----------
   // 标题：作业开始
   // 含义：将 #MainStep.S1 AND NOT (#MainStep.S2) 赋给 "DB1900_Communication_PC".Send.WorkStart
   "DB1900_Communication_PC".Send.WorkStart := #MainStep.S1 AND NOT (#MainStep.S2);
   // 含义：条件 #MainStep.S1 AND NOT (#MainStep.S2) 成立时，将 50 传送到 "DB1080_Component".Robot.CTRL_IN.RobotSpeed
   IF #MainStep.S1 AND NOT (#MainStep.S2) THEN
       "DB1080_Component".Robot.CTRL_IN.RobotSpeed := 50;
   END_IF;
   // 含义：将 (#MainStep.S1 AND "DB1900_Communication_PC".Recv.WorkStart) OR (#MainStep.S1 AND #MainStep.S2) 赋给 #MainStep.S2
   #MainStep.S2 := (#MainStep.S1 AND "DB1900_Communication_PC".Recv.WorkStart) OR (#MainStep.S1 AND #MainStep.S2);

   // ---------- 网络 7 ----------
   // 标题：参数写入
   // 含义：条件 #MainStep.S2 AND NOT (#MainStep.S3) 成立时，将 TRUE 传送到 "DB1081_ValveCall".ST01.Z08.RetAuto
   IF #MainStep.S2 AND NOT (#MainStep.S3) THEN
       "DB1081_ValveCall".ST01.Z08.RetAuto := TRUE;
   END_IF;
   // 含义：当 #MainStep.S2 为 TRUE 时置位 #MainStep.S3，否则复位（触点→线圈）
   IF #MainStep.S2 THEN
       #MainStep.S3 := TRUE;
   ELSE
       #MainStep.S3 := FALSE;
   END_IF;

   // ---------- 网络 8 ----------
   // 标题：S5 判断夹爪  S14更换夹爪
   // 含义：将 ((((#MainStep.S3 AND NOT (#EdgeDetc.Pulse[0])) AND NOT (#EdgeDetc.Pulse[0])) AND "DB720_KuKa_MainCtrl".Aux.ToolAtPosTimer.Q) OR (((#MainStep.S3 AND NOT (#EdgeDetc.Pulse[0])) AND NOT (#EdgeDetc.Pulse[0])) AND #MainStep.S5)) AND NOT (#MainStep.S14) 赋给 #MainStep.S5
   #MainStep.S5 := ((((#MainStep.S3 AND NOT (#EdgeDetc.Pulse[0])) AND NOT (#EdgeDetc.Pulse[0])) AND "DB720_KuKa_MainCtrl".Aux.ToolAtPosTimer.Q) OR (((#MainStep.S3 AND NOT (#EdgeDetc.Pulse[0])) AND NOT (#EdgeDetc.Pulse[0])) AND #MainStep.S5)) AND NOT (#MainStep.S14);
   // 含义：将 ((((#MainStep.S3 AND NOT (#EdgeDetc.Pulse[0])) AND NOT (#EdgeDetc.Pulse[0])) AND "DB720_KuKa_MainCtrl".Aux.ToolNotAtPosTimer.Q) OR (((#MainStep.S3 AND NOT (#EdgeDetc.Pulse[0])) AND NOT (#EdgeDetc.Pulse[0])) AND #MainStep.S14)) AND NOT (#MainStep.S5) 赋给 #MainStep.S14
   #MainStep.S14 := ((((#MainStep.S3 AND NOT (#EdgeDetc.Pulse[0])) AND NOT (#EdgeDetc.Pulse[0])) AND "DB720_KuKa_MainCtrl".Aux.ToolNotAtPosTimer.Q) OR (((#MainStep.S3 AND NOT (#EdgeDetc.Pulse[0])) AND NOT (#EdgeDetc.Pulse[0])) AND #MainStep.S14)) AND NOT (#MainStep.S5);

   // ---------- 网络 9 ----------
   // 标题：请求上位机参数录入...
   // 含义：条件 #MainStep.S5 AND NOT (#MainStep.S7) 成立时，将 TRUE 传送到 "DB1081_ValveCall".ST01.Z08.ExtAuto
   IF #MainStep.S5 AND NOT (#MainStep.S7) THEN
       "DB1081_ValveCall".ST01.Z08.ExtAuto := TRUE;
   END_IF;
   // 含义：将 #MainStep.S5 AND NOT (#MainStep.S7) 赋给 "DB1146_PromptFree".Public.AskPcData
   "DB1146_PromptFree".Public.AskPcData := #MainStep.S5 AND NOT (#MainStep.S7);
   // 含义：将 (((#MainStep.S5 AND "DB1900_Communication_PC".Recv.ParaWriteDone) AND NOT ("DB1080_Component".Robot.Status.Busy)) AND "DB1081_ValveCall".ST01.Z08.ExtPos) OR (#MainStep.S5 AND #MainStep.S7) 赋给 #MainStep.S7
   #MainStep.S7 := (((#MainStep.S5 AND "DB1900_Communication_PC".Recv.ParaWriteDone) AND NOT ("DB1080_Component".Robot.Status.Busy)) AND "DB1081_ValveCall".ST01.Z08.ExtPos) OR (#MainStep.S5 AND #MainStep.S7);
   // 含义：调用计数器实例 "Timer_ParaWriteOuttime".TON（上升沿计数，当前值写入 CV）
   "Timer_ParaWriteOuttime".TON(IN := (#MainStep.S5 AND NOT (#MainStep.S7)) AND NOT ("DB1900_Communication_PC".Recv.ParaWriteDone),
                                PT := t#5s);
   // 含义：条件 "Timer_ParaWriteOuttime".Q 成立时，将 TRUE 传送到 #MainStep.ErrEnd
   IF "Timer_ParaWriteOuttime".Q THEN
       #MainStep.ErrEnd := TRUE;
   END_IF;
   // 含义：条件 "Timer_ParaWriteOuttime".Q 成立时，将 FALSE 传送到 "DB1900_Communication_PC".Send.PowerOff
   IF "Timer_ParaWriteOuttime".Q THEN
       "DB1900_Communication_PC".Send.PowerOff := FALSE;
   END_IF;
   // 含义：条件 "Timer_ParaWriteOuttime".Q 成立时，将 TRUE 传送到 "DB1147_PromptStartNotPmt".Public.ParaWiriteOuttime
   IF "Timer_ParaWriteOuttime".Q THEN
       "DB1147_PromptStartNotPmt".Public.ParaWiriteOuttime := TRUE;
   END_IF;

   // ---------- 网络 10 ----------
   // 标题：钻孔方向
   // 含义：条件 (#MainStep.S7 AND NOT (#MainStep.S8)) AND "DB1900_Communication_PC".Para.DrillDirection1 成立时，将 1 传送到 "DB1042_Timer".DrillDirectionCurrent
   IF (#MainStep.S7 AND NOT (#MainStep.S8)) AND "DB1900_Communication_PC".Para.DrillDirection1 THEN
       "DB1042_Timer".DrillDirectionCurrent := 1;
   END_IF;
   // 含义：条件 (#MainStep.S7 AND NOT (#MainStep.S8)) AND "DB1900_Communication_PC".Para.DrillDirection2 成立时，将 2 传送到 "DB1042_Timer".DrillDirectionCurrent
   IF (#MainStep.S7 AND NOT (#MainStep.S8)) AND "DB1900_Communication_PC".Para.DrillDirection2 THEN
       "DB1042_Timer".DrillDirectionCurrent := 2;
   END_IF;
   // 含义：条件 (#MainStep.S7 AND NOT (#MainStep.S8)) AND "DB1900_Communication_PC".Para.DrillDirection3 成立时，将 3 传送到 "DB1042_Timer".DrillDirectionCurrent
   IF (#MainStep.S7 AND NOT (#MainStep.S8)) AND "DB1900_Communication_PC".Para.DrillDirection3 THEN
       "DB1042_Timer".DrillDirectionCurrent := 3;
   END_IF;
   // 含义：条件 ((#MainStep.S7 AND NOT (#MainStep.S8)) AND ("DB1042_Timer".DrillDirectionMemory <> "DB1042_Timer".DrillDirectionCurrent)) 成立时，将 0 传送到 #Aux.HoleNo
   IF ((#MainStep.S7 AND NOT (#MainStep.S8)) AND ("DB1042_Timer".DrillDirectionMemory <> "DB1042_Timer".DrillDirectionCurrent)) THEN
       #Aux.HoleNo := 0;
   END_IF;
   // 含义：将 ((#MainStep.S7 AND (#Aux.HoleNo = 0))) OR ((#MainStep.S7 AND ("DB1042_Timer".DrillDirectionMemory = "DB1042_Timer".DrillDirectionCurrent))) OR (#MainStep.S7 AND #MainStep.S8) 赋给 #MainStep.S8
   #MainStep.S8 := ((#MainStep.S7 AND (#Aux.HoleNo = 0))) OR ((#MainStep.S7 AND ("DB1042_Timer".DrillDirectionMemory = "DB1042_Timer".DrillDirectionCurrent))) OR (#MainStep.S7 AND #MainStep.S8);

   // ---------- 网络 11 ----------
   // 标题：参数写入
   // 含义：条件 #MainStep.S8 AND NOT (#MainStep.S9) 成立时，将 TRUE 传送到 "DB1081_ValveCall".ST01.Z08.ExtAuto
   IF #MainStep.S8 AND NOT (#MainStep.S9) THEN
       "DB1081_ValveCall".ST01.Z08.ExtAuto := TRUE;
   END_IF;
   // 含义：条件 #MainStep.S8 AND NOT (#MainStep.S9) 成立时，将 TRUE 传送到 "DB1080_Component".Robot.Cmd.Auto.GoHome
   IF #MainStep.S8 AND NOT (#MainStep.S9) THEN
       "DB1080_Component".Robot.Cmd.Auto.GoHome := TRUE;
   END_IF;
   // 含义：条件 (#MainStep.S8 AND NOT (#MainStep.S9)) AND "DB1900_Communication_PC".Para.DrillDirection1 成立时，将 1 传送到 "DB1042_Timer".DrillDirectionMemory
   IF (#MainStep.S8 AND NOT (#MainStep.S9)) AND "DB1900_Communication_PC".Para.DrillDirection1 THEN
       "DB1042_Timer".DrillDirectionMemory := 1;
   END_IF;
   // 含义：条件 (#MainStep.S8 AND NOT (#MainStep.S9)) AND "DB1900_Communication_PC".Para.DrillDirection2 成立时，将 2 传送到 "DB1042_Timer".DrillDirectionMemory
   IF (#MainStep.S8 AND NOT (#MainStep.S9)) AND "DB1900_Communication_PC".Para.DrillDirection2 THEN
       "DB1042_Timer".DrillDirectionMemory := 2;
   END_IF;
   // 含义：条件 (#MainStep.S8 AND NOT (#MainStep.S9)) AND "DB1900_Communication_PC".Para.DrillDirection3 成立时，将 3 传送到 "DB1042_Timer".DrillDirectionMemory
   IF (#MainStep.S8 AND NOT (#MainStep.S9)) AND "DB1900_Communication_PC".Para.DrillDirection3 THEN
       "DB1042_Timer".DrillDirectionMemory := 3;
   END_IF;
   // 含义：将 (#MainStep.S8 AND "DB1080_Component".Robot.Status.HomePos) OR (#MainStep.S8 AND #MainStep.S9) 赋给 #MainStep.S9
   #MainStep.S9 := (#MainStep.S8 AND "DB1080_Component".Robot.Status.HomePos) OR (#MainStep.S8 AND #MainStep.S9);

   // ---------- 网络 12 ----------
   // 标题：JUMP[4]需要换型  S20不需要
   // 注释：钻孔时，仅有S20线圈导通
   // 含义：将 ((((#MainStep.S9 AND NOT (#EdgeDetc.Pulse[0])) AND NOT (#MainStep.S20)) AND NOT (#EdgeDetc.Pulse[0])) AND ("DB1900_Communication_PC".Para.IOFixtureNo <> "DB1080_Component".IOFixtureIID.TP_CurFixtureID)) 赋给 "DB1148_PromptBeeper".Public.IoToolNoCompErr
   "DB1148_PromptBeeper".Public.IoToolNoCompErr := ((((#MainStep.S9 AND NOT (#EdgeDetc.Pulse[0])) AND NOT (#MainStep.S20)) AND NOT (#EdgeDetc.Pulse[0])) AND ("DB1900_Communication_PC".Para.IOFixtureNo <> "DB1080_Component".IOFixtureIID.TP_CurFixtureID));
   // 含义：将 ((((#MainStep.S9 AND NOT (#EdgeDetc.Pulse[0])) AND NOT (#MainStep.S20)) AND NOT (#EdgeDetc.Pulse[0])) AND ("DB1900_Communication_PC".Para.PowerFixtureNo <> "DB1080_Component".PowerFixtureID.TP_CurFixtureID)) 赋给 "DB1148_PromptBeeper".Public.PowerToolNoCompErr
   "DB1148_PromptBeeper".Public.PowerToolNoCompErr := ((((#MainStep.S9 AND NOT (#EdgeDetc.Pulse[0])) AND NOT (#MainStep.S20)) AND NOT (#EdgeDetc.Pulse[0])) AND ("DB1900_Communication_PC".Para.PowerFixtureNo <> "DB1080_Component".PowerFixtureID.TP_CurFixtureID));
   // 含义：将 (((((((#MainStep.S9 AND NOT (#EdgeDetc.Pulse[0])) AND "DB720_KuKa_MainCtrl".Aux.ToolAtPosTimer.Q) AND ("DB1900_Communication_PC".Para.IOFixtureNo = "DB1080_Component".IOFixtureIID.TP_CurFixtureID))) AND ("DB1900_Communication_PC".Para.PowerFixtureNo = "DB1080_Component".PowerFixtureID.TP_CurFixtureID))) OR ((#MainStep.S9 AND NOT (#EdgeDetc.Pulse[0])) AND #MainStep.S20)) AND NOT (#EdgeDetc.Pulse[0]) 赋给 #MainStep.S20
   #MainStep.S20 := (((((((#MainStep.S9 AND NOT (#EdgeDetc.Pulse[0])) AND "DB720_KuKa_MainCtrl".Aux.ToolAtPosTimer.Q) AND ("DB1900_Communication_PC".Para.IOFixtureNo = "DB1080_Component".IOFixtureIID.TP_CurFixtureID))) AND ("DB1900_Communication_PC".Para.PowerFixtureNo = "DB1080_Component".PowerFixtureID.TP_CurFixtureID))) OR ((#MainStep.S9 AND NOT (#EdgeDetc.Pulse[0])) AND #MainStep.S20)) AND NOT (#EdgeDetc.Pulse[0]);
   // 含义：将 ((((#MainStep.S9 AND NOT (#EdgeDetc.Pulse[0])) AND "ErrRst_M") AND "DB1148_PromptBeeper".Public.IoToolNoCompErr) OR (((#MainStep.S9 AND NOT (#EdgeDetc.Pulse[0])) AND "ErrRst_M") AND "DB1148_PromptBeeper".Public.PowerToolNoCompErr) OR ((#MainStep.S9 AND NOT (#EdgeDetc.Pulse[0])) AND #EdgeDetc.Pulse[0])) AND NOT (#MainStep.S20) 赋给 #EdgeDetc.Pulse[0]
   #EdgeDetc.Pulse[0] := ((((#MainStep.S9 AND NOT (#EdgeDetc.Pulse[0])) AND "ErrRst_M") AND "DB1148_PromptBeeper".Public.IoToolNoCompErr) OR (((#MainStep.S9 AND NOT (#EdgeDetc.Pulse[0])) AND "ErrRst_M") AND "DB1148_PromptBeeper".Public.PowerToolNoCompErr) OR ((#MainStep.S9 AND NOT (#EdgeDetc.Pulse[0])) AND #EdgeDetc.Pulse[0])) AND NOT (#MainStep.S20);

   // ---------- 网络 13 ----------
   // 标题：机器人状态
   // 注释：钻孔时，S22导通并自保持
   // 含义：将 (((#MainStep.S20 AND NOT (#RobotAutoStep.Status.Running)) AND NOT (#RobotAutoStep.CheckBitStatus.TaskDone)) AND NOT (#RobotAutoStep.DrillStatus.TaskDone)) OR (#MainStep.S20 AND #MainStep.S22) 赋给 #MainStep.S22
   #MainStep.S22 := (((#MainStep.S20 AND NOT (#RobotAutoStep.Status.Running)) AND NOT (#RobotAutoStep.CheckBitStatus.TaskDone)) AND NOT (#RobotAutoStep.DrillStatus.TaskDone)) OR (#MainStep.S20 AND #MainStep.S22);
   // 含义：条件 #MainStep.S20 AND NOT (#MainStep.S22) 成立时，将 FALSE 传送到 #RobotAutoStep.CheckBitStatus.TaskDone
   IF #MainStep.S20 AND NOT (#MainStep.S22) THEN
       #RobotAutoStep.CheckBitStatus.TaskDone := FALSE;
   END_IF;
   // 含义：条件 #MainStep.S20 AND NOT (#MainStep.S22) 成立时，将 FALSE 传送到 #RobotAutoStep.DrillStatus.TaskDone
   IF #MainStep.S20 AND NOT (#MainStep.S22) THEN
       #RobotAutoStep.DrillStatus.TaskDone := FALSE;
   END_IF;

   // ---------- 网络 14 ----------
   // 标题：S25 第一颗螺丝先校准   S27不需要校准
   // 含义：将 (((#MainStep.S22 AND #Status.FirstStart) AND NOT ("DB1900_Communication_PC".Recv.DrillStart)) OR (#MainStep.S22 AND #MainStep.S25)) AND NOT (#MainStep.S27) 赋给 #MainStep.S25
   #MainStep.S25 := (((#MainStep.S22 AND #Status.FirstStart) AND NOT ("DB1900_Communication_PC".Recv.DrillStart)) OR (#MainStep.S22 AND #MainStep.S25)) AND NOT (#MainStep.S27);
   // 含义：将 ((#MainStep.S22 AND NOT (#MainStep.S25)) AND "DB1900_Communication_PC".Recv.DrillStart) OR (#MainStep.S22 AND #MainStep.S27) 赋给 #MainStep.S27
   #MainStep.S27 := ((#MainStep.S22 AND NOT (#MainStep.S25)) AND "DB1900_Communication_PC".Recv.DrillStart) OR (#MainStep.S22 AND #MainStep.S27);

   // ---------- 网络 15 ----------
   // 标题：更换电锤完成
   // 含义：将 (#MainStep.S25 AND NOT (#MainStep.S30)) OR ((((#MainStep.S1 AND NOT (#MainStep.S2)) AND NOT ("DB720_KuKa_MainCtrl".Aux.ToolAtPos)) AND NOT ("DB1900_Communication_PC".Recv.DrillStart)) AND NOT ("DB720_KuKa_MainCtrl".StatusIn.do_ChgGrp_Don)) OR ((((NOT ("DB1042_Timer".FirstStart) AND "DB1900_Communication_PC".Send.DrillStart) AND NOT ("DB1900_Communication_PC".Recv.DrillStart)) AND ("DB720_KuKa_MainCtrl".CmdOut.gi_ToolTypeNo <> 2))) 赋给 "DB1900_Communication_PC".Send.ChangeToolDone
   "DB1900_Communication_PC".Send.ChangeToolDone := (#MainStep.S25 AND NOT (#MainStep.S30)) OR ((((#MainStep.S1 AND NOT (#MainStep.S2)) AND NOT ("DB720_KuKa_MainCtrl".Aux.ToolAtPos)) AND NOT ("DB1900_Communication_PC".Recv.DrillStart)) AND NOT ("DB720_KuKa_MainCtrl".StatusIn.do_ChgGrp_Don)) OR ((((NOT ("DB1042_Timer".FirstStart) AND "DB1900_Communication_PC".Send.DrillStart) AND NOT ("DB1900_Communication_PC".Recv.DrillStart)) AND ("DB720_KuKa_MainCtrl".CmdOut.gi_ToolTypeNo <> 2)));

   // ---------- 网络 16 ----------
   // 标题：校验
   // 含义：条件 (#MainStep.S25 AND NOT (#MainStep.S26)) AND "DB1900_Communication_PC".Recv.Z05RetTPPB 成立时，将 TRUE 传送到 #RobotAutoStep.Cmd.Auto.CheckBit
   IF (#MainStep.S25 AND NOT (#MainStep.S26)) AND "DB1900_Communication_PC".Recv.Z05RetTPPB THEN
       #RobotAutoStep.Cmd.Auto.CheckBit := TRUE;
   END_IF;
   // 含义：条件 #MainStep.S25 AND NOT (#MainStep.S26) 成立时，将 TRUE 传送到 "DB1042_Timer".FirstStart
   IF #MainStep.S25 AND NOT (#MainStep.S26) THEN
       "DB1042_Timer".FirstStart := TRUE;
   END_IF;
   // 含义：将 ((#MainStep.S25 AND #RobotAutoStep.CheckBitStatus.TaskDone) AND #RobotAutoStep.CheckBitStatus.TaskIO) OR (#MainStep.S25 AND #MainStep.S26) 赋给 #MainStep.S26
   #MainStep.S26 := ((#MainStep.S25 AND #RobotAutoStep.CheckBitStatus.TaskDone) AND #RobotAutoStep.CheckBitStatus.TaskIO) OR (#MainStep.S25 AND #MainStep.S26);
   // 含义：条件 (#MainStep.S25 AND #RobotAutoStep.CheckBitStatus.TaskDone) AND #RobotAutoStep.CheckBitStatus.TaskNIO 成立时，将 TRUE 传送到 #MainStep.ErrEnd
   IF (#MainStep.S25 AND #RobotAutoStep.CheckBitStatus.TaskDone) AND #RobotAutoStep.CheckBitStatus.TaskNIO THEN
       #MainStep.ErrEnd := TRUE;
   END_IF;

   // ---------- 网络 17 ----------
   // 标题：请求热机
   // 含义：将 #MainStep.S26 AND NOT (#MainStep.S30) 赋给 "DB1900_Communication_PC".Send.ReqHeatMachine
   "DB1900_Communication_PC".Send.ReqHeatMachine := #MainStep.S26 AND NOT (#MainStep.S30);
   // 含义：将 #MainStep.S26 AND NOT (#MainStep.S30) 赋给 "DB1146_PromptFree".ST01.HeatMachin
   "DB1146_PromptFree".ST01.HeatMachin := #MainStep.S26 AND NOT (#MainStep.S30);
   // 含义：条件 (#MainStep.S26 AND NOT (#MainStep.S30)) AND NOT (TRUE) 成立时，将 TRUE 传送到 "DB1081_ValveCall".ST01.Z05.ExtAuto
   IF (#MainStep.S26 AND NOT (#MainStep.S30)) AND NOT (TRUE) THEN
       "DB1081_ValveCall".ST01.Z05.ExtAuto := TRUE;
   END_IF;
   // 含义：将 (#MainStep.S26 AND "DB1900_Communication_PC".Recv.ResHeatMachin) OR (#MainStep.S26 AND #MainStep.S30) 赋给 #MainStep.S30
   #MainStep.S30 := (#MainStep.S26 AND "DB1900_Communication_PC".Recv.ResHeatMachin) OR (#MainStep.S26 AND #MainStep.S30);

   // ---------- 网络 18 ----------
   // 标题：打孔流程启动
   // 注释：流程边界问题：规程结束时刚好打完一个孔，要去打下一个孔，Recv.DrillStart信号立即为False, MainStep32未接通，之后的流程不通，机器人停在水泥块表面 ，工具未断电。更改：将JUMP[0]信号并入条件
   // 含义：将 (((((((((((#MainStep.S30 OR #MainStep.S27) AND NOT (#EdgeDetc.Pulse[0])) AND NOT (#RobotAutoStep.Status.Running)) AND NOT (#RobotAutoStep.DrillStatus.TaskDone)) AND NOT ("DB1080_Component".Robot.Status.Busy)) AND "DB1900_Communication_PC".Recv.DrillStart) OR ((((((((#MainStep.S30 OR #MainStep.S27) AND NOT (#EdgeDetc.Pulse[0])) AND NOT (#RobotAutoStep.Status.Running)) AND NOT (#RobotAutoStep.DrillStatus.TaskDone)) AND NOT ("DB1080_Component".Robot.Status.Busy)) AND NOT ("DB1900_Communication_PC".Recv.DrillStart)) AND "DB1900_Communication_PC".Send.DrillRunning) AND NOT (#EdgeDetc.Pulse[0]))) AND ("DB1900_Communication_PC".Para.IOFixtureNo = "DB1080_Component".IOFixtureIID.TP_CurFixtureID))) AND ("DB1900_Communication_PC".Para.PowerFixtureNo = "DB1080_Component".PowerFixtureID.TP_CurFixtureID))) OR (((#MainStep.S30 OR #MainStep.S27) AND NOT (#EdgeDetc.Pulse[0])) AND #MainStep.S32) 赋给 #MainStep.S32
   #MainStep.S32 := (((((((((((#MainStep.S30 OR #MainStep.S27) AND NOT (#EdgeDetc.Pulse[0])) AND NOT (#RobotAutoStep.Status.Running)) AND NOT (#RobotAutoStep.DrillStatus.TaskDone)) AND NOT ("DB1080_Component".Robot.Status.Busy)) AND "DB1900_Communication_PC".Recv.DrillStart) OR ((((((((#MainStep.S30 OR #MainStep.S27) AND NOT (#EdgeDetc.Pulse[0])) AND NOT (#RobotAutoStep.Status.Running)) AND NOT (#RobotAutoStep.DrillStatus.TaskDone)) AND NOT ("DB1080_Component".Robot.Status.Busy)) AND NOT ("DB1900_Communication_PC".Recv.DrillStart)) AND "DB1900_Communication_PC".Send.DrillRunning) AND NOT (#EdgeDetc.Pulse[0]))) AND ("DB1900_Communication_PC".Para.IOFixtureNo = "DB1080_Component".IOFixtureIID.TP_CurFixtureID))) AND ("DB1900_Communication_PC".Para.PowerFixtureNo = "DB1080_Component".PowerFixtureID.TP_CurFixtureID))) OR (((#MainStep.S30 OR #MainStep.S27) AND NOT (#EdgeDetc.Pulse[0])) AND #MainStep.S32);
   // 含义：将 (((((#MainStep.S30 OR #MainStep.S27) AND NOT (#EdgeDetc.Pulse[0])) AND ("DB1900_Communication_PC".Para.IOFixtureNo <> "DB1080_Component".IOFixtureIID.TP_CurFixtureID))) OR ((((#MainStep.S30 OR #MainStep.S27) AND NOT (#EdgeDetc.Pulse[0])) AND ("DB1900_Communication_PC".Para.PowerFixtureNo <> "DB1080_Component".PowerFixtureID.TP_CurFixtureID)))) AND NOT (#MainStep.S32) 赋给 #EdgeDetc.Pulse[0]
   #EdgeDetc.Pulse[0] := (((((#MainStep.S30 OR #MainStep.S27) AND NOT (#EdgeDetc.Pulse[0])) AND ("DB1900_Communication_PC".Para.IOFixtureNo <> "DB1080_Component".IOFixtureIID.TP_CurFixtureID))) OR ((((#MainStep.S30 OR #MainStep.S27) AND NOT (#EdgeDetc.Pulse[0])) AND ("DB1900_Communication_PC".Para.PowerFixtureNo <> "DB1080_Component".PowerFixtureID.TP_CurFixtureID)))) AND NOT (#MainStep.S32);
   // 含义：将 ((#MainStep.S30 OR #MainStep.S27 OR (#MainStep.S22 AND NOT (#MainStep.S25))) AND NOT (#EdgeDetc.Pulse[0])) AND NOT (#MainStep.S32) 赋给 "DB1900_Communication_PC".Send.DrillStart
   "DB1900_Communication_PC".Send.DrillStart := ((#MainStep.S30 OR #MainStep.S27 OR (#MainStep.S22 AND NOT (#MainStep.S25))) AND NOT (#EdgeDetc.Pulse[0])) AND NOT (#MainStep.S32);
   // 含义：条件 ((#MainStep.S30 OR #MainStep.S27 OR (#MainStep.S22 AND NOT (#MainStep.S25))) AND NOT (#EdgeDetc.Pulse[0])) AND NOT (#MainStep.S32) 成立时，将 FALSE 传送到 #RobotAutoStep.DrillStatus.TaskDone
   IF ((#MainStep.S30 OR #MainStep.S27 OR (#MainStep.S22 AND NOT (#MainStep.S25))) AND NOT (#EdgeDetc.Pulse[0])) AND NOT (#MainStep.S32) THEN
       #RobotAutoStep.DrillStatus.TaskDone := FALSE;
   END_IF;

   // ---------- 网络 19 ----------
   // 含义：当 #MainStep.S32 为 TRUE 时置位 #MainStep.S34，否则复位（触点→线圈）
   IF #MainStep.S32 THEN
       #MainStep.S34 := TRUE;
   ELSE
       #MainStep.S34 := FALSE;
   END_IF;

   // ---------- 网络 20 ----------
   // 标题：钻孔
   // 含义：条件 #MainStep.S34 AND NOT (#MainStep.S35) 成立时，将 TRUE 传送到 #RobotAutoStep.Cmd.Auto.Drill
   IF #MainStep.S34 AND NOT (#MainStep.S35) THEN
       #RobotAutoStep.Cmd.Auto.Drill := TRUE;
   END_IF;
   // 含义：条件 #MainStep.S34 AND NOT (#MainStep.S35) 成立时，将 TRUE 传送到 "DB1042_Timer".DrillMemory
   IF #MainStep.S34 AND NOT (#MainStep.S35) THEN
       "DB1042_Timer".DrillMemory := TRUE;
   END_IF;
   // 含义：条件 #MainStep.S34 AND NOT (#MainStep.S35) 成立时，将 TRUE 传送到 "DB1900_Communication_PC".Send.DrillRunning
   IF #MainStep.S34 AND NOT (#MainStep.S35) THEN
       "DB1900_Communication_PC".Send.DrillRunning := TRUE;
   END_IF;
   // 含义：条件 #MainStep.S34 AND NOT (#MainStep.S35) 成立时，将 FALSE 传送到 #Status.FirstStart
   IF #MainStep.S34 AND NOT (#MainStep.S35) THEN
       #Status.FirstStart := FALSE;
   END_IF;
   // 含义：条件 (((#MainStep.S34 AND NOT (#MainStep.S35)) AND #HorDrillAutoStep.HorDrillStep.StopDrill_Ack) OR ((#MainStep.S34 AND NOT (#MainStep.S35)) AND #DownDrillAutoStep.DownDrillStep.StopDrill_Ack)) AND NOT (#EdgeDetc.Pulse[0]) 成立时，将 (#Aux.HoleNo + 1) 传送到 #Aux.HoleNo
   IF (((#MainStep.S34 AND NOT (#MainStep.S35)) AND #HorDrillAutoStep.HorDrillStep.StopDrill_Ack) OR ((#MainStep.S34 AND NOT (#MainStep.S35)) AND #DownDrillAutoStep.DownDrillStep.StopDrill_Ack)) AND NOT (#EdgeDetc.Pulse[0]) THEN
       #Aux.HoleNo := (#Aux.HoleNo + 1);
   END_IF;
   // 含义：将 ((#MainStep.S34 AND NOT (#MainStep.S35)) AND #HorDrillAutoStep.HorDrillStep.StopDrill_Ack) OR ((#MainStep.S34 AND NOT (#MainStep.S35)) AND #DownDrillAutoStep.DownDrillStep.StopDrill_Ack) 赋给 #EdgeDetc.Pulse[0]
   #EdgeDetc.Pulse[0] := ((#MainStep.S34 AND NOT (#MainStep.S35)) AND #HorDrillAutoStep.HorDrillStep.StopDrill_Ack) OR ((#MainStep.S34 AND NOT (#MainStep.S35)) AND #DownDrillAutoStep.DownDrillStep.StopDrill_Ack);
   // 含义：将 ((#MainStep.S34 AND #RobotAutoStep.DrillStatus.TaskDone) AND #RobotAutoStep.DrillStatus.TaskIO) OR (#MainStep.S34 AND #MainStep.S35) 赋给 #MainStep.S35
   #MainStep.S35 := ((#MainStep.S34 AND #RobotAutoStep.DrillStatus.TaskDone) AND #RobotAutoStep.DrillStatus.TaskIO) OR (#MainStep.S34 AND #MainStep.S35);
   // 含义：条件 (#MainStep.S34 AND #RobotAutoStep.DrillStatus.TaskDone) AND #RobotAutoStep.DrillStatus.TaskNIO 成立时，将 TRUE 传送到 "DB1081_ValveCall".ST01.Z05.RetAuto
   IF (#MainStep.S34 AND #RobotAutoStep.DrillStatus.TaskDone) AND #RobotAutoStep.DrillStatus.TaskNIO THEN
       "DB1081_ValveCall".ST01.Z05.RetAuto := TRUE;
   END_IF;
   // 含义：条件 (#MainStep.S34 AND #RobotAutoStep.DrillStatus.TaskDone) AND #RobotAutoStep.DrillStatus.TaskNIO 成立时，将 TRUE 传送到 #MainStep.ErrEnd
   IF (#MainStep.S34 AND #RobotAutoStep.DrillStatus.TaskDone) AND #RobotAutoStep.DrillStatus.TaskNIO THEN
       #MainStep.ErrEnd := TRUE;
   END_IF;
   // 含义：条件 ((#MainStep.S34 AND #RobotAutoStep.DrillStatus.TaskDone) AND #RobotAutoStep.DrillStatus.TaskNIO) AND NOT ("DB1900_Communication_PC".Recv.PowerOff) 成立时，将 TRUE 传送到 "DB1900_Communication_PC".Send.PowerOff
   IF ((#MainStep.S34 AND #RobotAutoStep.DrillStatus.TaskDone) AND #RobotAutoStep.DrillStatus.TaskNIO) AND NOT ("DB1900_Communication_PC".Recv.PowerOff) THEN
       "DB1900_Communication_PC".Send.PowerOff := TRUE;
   END_IF;

   // ---------- 网络 21 ----------
   // 标题：用作打击记忆，回原点开枪
   // 含义：条件 #MainStep.S35 AND NOT (#MainStep.S37) 成立时，将 FALSE 传送到 "DB1042_Timer".DrillMemory
   IF #MainStep.S35 AND NOT (#MainStep.S37) THEN
       "DB1042_Timer".DrillMemory := FALSE;
   END_IF;
   // 含义：当 #MainStep.S35 为 TRUE 时置位 #MainStep.S37，否则复位（触点→线圈）
   IF #MainStep.S35 THEN
       #MainStep.S37 := TRUE;
   ELSE
       #MainStep.S37 := FALSE;
   END_IF;

   // ---------- 网络 22 ----------
   // 标题：打孔中
   // 注释：#EdgeDetc.JUMP[8] : Robot Go to Home Position then Put Gripper in Station  when  Intermedirate Test  End
   // 含义：将 #MainStep.S37 AND NOT ("DB1900_Communication_PC".Recv.DrillStart) 赋给 #EdgeDetc.Pulse[0]
   #EdgeDetc.Pulse[0] := #MainStep.S37 AND NOT ("DB1900_Communication_PC".Recv.DrillStart);
   // 含义：条件 #MainStep.S37 AND NOT ("DB1900_Communication_PC".Recv.DrillStart) 成立时，将 FALSE 传送到 "DB1900_Communication_PC".Send.DrillRunning
   IF #MainStep.S37 AND NOT ("DB1900_Communication_PC".Recv.DrillStart) THEN
       "DB1900_Communication_PC".Send.DrillRunning := FALSE;
   END_IF;
   // 含义：将 #MainStep.S37 AND "DB1900_Communication_PC".Recv.WorkDone 赋给 "DB1900_Communication_PC".Send.WorkDone
   "DB1900_Communication_PC".Send.WorkDone := #MainStep.S37 AND "DB1900_Communication_PC".Recv.WorkDone;

   // ---------- 网络 23 ----------
   // 标题：换枪和继续打孔 依据上位机命令 50结束 40换枪  JUMP[0]继续打孔, 57岩芯敲击
   // 注释：按打孔数结束完全由上位机来控制
   // 含义：将 (#MainStep.S37 AND "DB1900_Communication_PC".Recv.DrillStart) AND NOT (#MainStep.S40) 赋给 #EdgeDetc.Pulse[0]
   #EdgeDetc.Pulse[0] := (#MainStep.S37 AND "DB1900_Communication_PC".Recv.DrillStart) AND NOT (#MainStep.S40);
   // 含义：条件 (#MainStep.S37 AND "DB1900_Communication_PC".Recv.DrillStart) AND NOT (#MainStep.S40) 成立时，将 FALSE 传送到 #RobotAutoStep.DrillStatus.TaskDone
   IF (#MainStep.S37 AND "DB1900_Communication_PC".Recv.DrillStart) AND NOT (#MainStep.S40) THEN
       #RobotAutoStep.DrillStatus.TaskDone := FALSE;
   END_IF;
   // 含义：将 ((((((#MainStep.S37 AND NOT ("DB1900_Communication_PC".Recv.DrillStart)) AND NOT ("DB1900_Communication_PC".Recv.ChangeTool)) AND "DB1900_Communication_PC".Recv.WorkDone) OR (((#MainStep.S37 AND NOT ("DB1900_Communication_PC".Recv.DrillStart)) AND NOT ("DB1900_Communication_PC".Recv.ChangeTool)) AND NOT ("DB1900_Communication_PC".Recv.WorkStart))) AND NOT ("DB1900_Communication_PC".Para.ControlMode)) OR ((((((#MainStep.S37 AND NOT ("DB1900_Communication_PC".Recv.DrillStart)) AND NOT ("DB1900_Communication_PC".Recv.ChangeTool)) AND NOT (TRUE)) AND (#Aux.HoleNo >= "DB1900_Communication_PC".Para.HoleNum))) AND "DB1900_Communication_PC".Para.ControlMode) OR (#MainStep.S37 AND #MainStep.S50)) AND NOT (#MainStep.S40) 赋给 #MainStep.S50
   #MainStep.S50 := ((((((#MainStep.S37 AND NOT ("DB1900_Communication_PC".Recv.DrillStart)) AND NOT ("DB1900_Communication_PC".Recv.ChangeTool)) AND "DB1900_Communication_PC".Recv.WorkDone) OR (((#MainStep.S37 AND NOT ("DB1900_Communication_PC".Recv.DrillStart)) AND NOT ("DB1900_Communication_PC".Recv.ChangeTool)) AND NOT ("DB1900_Communication_PC".Recv.WorkStart))) AND NOT ("DB1900_Communication_PC".Para.ControlMode)) OR ((((((#MainStep.S37 AND NOT ("DB1900_Communication_PC".Recv.DrillStart)) AND NOT ("DB1900_Communication_PC".Recv.ChangeTool)) AND NOT (TRUE)) AND (#Aux.HoleNo >= "DB1900_Communication_PC".Para.HoleNum))) AND "DB1900_Communication_PC".Para.ControlMode) OR (#MainStep.S37 AND #MainStep.S50)) AND NOT (#MainStep.S40);
   // 含义：将 (((#MainStep.S37 AND #EdgeDetc.Pulse[0]) OR (#MainStep.S37 AND #MainStep.S40)) AND NOT (#EdgeDetc.Pulse[0])) AND NOT (#MainStep.S50) 赋给 #MainStep.S40
   #MainStep.S40 := (((#MainStep.S37 AND #EdgeDetc.Pulse[0]) OR (#MainStep.S37 AND #MainStep.S40)) AND NOT (#EdgeDetc.Pulse[0])) AND NOT (#MainStep.S50);
   // 含义：将 ((#MainStep.S37 AND NOT (#MainStep.S40)) AND NOT (#MainStep.S50)) AND NOT (#EdgeDetc.Pulse[0]) 赋给 "DB1146_PromptFree".Public.WaitPcCommond
   "DB1146_PromptFree".Public.WaitPcCommond := ((#MainStep.S37 AND NOT (#MainStep.S40)) AND NOT (#MainStep.S50)) AND NOT (#EdgeDetc.Pulse[0]);

   // ---------- 网络 24 ----------
   // 标题：机器人状态
   // 含义：将 ((#MainStep.S40 OR #MainStep.S14 OR #EdgeDetc.Pulse[0]) AND NOT (#RobotAutoStep.Status.Running)) OR ((#MainStep.S40 OR #MainStep.S14 OR #EdgeDetc.Pulse[0]) AND #MainStep.S42) 赋给 #MainStep.S42
   #MainStep.S42 := ((#MainStep.S40 OR #MainStep.S14 OR #EdgeDetc.Pulse[0]) AND NOT (#RobotAutoStep.Status.Running)) OR ((#MainStep.S40 OR #MainStep.S14 OR #EdgeDetc.Pulse[0]) AND #MainStep.S42);

   // ---------- 网络 25 ----------
   // 含义：将 (#MainStep.S42 AND NOT ("DB1080_Component".Robot.Status.Busy)) OR (#MainStep.S42 AND #MainStep.S43) 赋给 #MainStep.S43
   #MainStep.S43 := (#MainStep.S42 AND NOT ("DB1080_Component".Robot.Status.Busy)) OR (#MainStep.S42 AND #MainStep.S43);

   // ---------- 网络 26 ----------
   // 标题：规程结束回原点
   // 含义：条件 (#MainStep.S43 AND NOT (#MainStep.S44)) AND "DB720_KuKa_MainCtrl".Aux.ToolAtPosTimer.Q 成立时，将 TRUE 传送到 "DB1080_Component".Robot.Cmd.Auto.GoHome
   IF (#MainStep.S43 AND NOT (#MainStep.S44)) AND "DB720_KuKa_MainCtrl".Aux.ToolAtPosTimer.Q THEN
       "DB1080_Component".Robot.Cmd.Auto.GoHome := TRUE;
   END_IF;
   // 含义：条件 #MainStep.S43 AND NOT (#MainStep.S44) 成立时，将 TRUE 传送到 "DB1081_ValveCall".ST01.Z08.RetAuto
   IF #MainStep.S43 AND NOT (#MainStep.S44) THEN
       "DB1081_ValveCall".ST01.Z08.RetAuto := TRUE;
   END_IF;
   // 含义：将 (#MainStep.S43 AND "DB1080_Component".Robot.Status.HomePos) OR (#MainStep.S43 AND #MainStep.S44) 赋给 #MainStep.S44
   #MainStep.S44 := (#MainStep.S43 AND "DB1080_Component".Robot.Status.HomePos) OR (#MainStep.S43 AND #MainStep.S44);

   // ---------- 网络 27 ----------
   // 含义：条件 ((((#MainStep.S44 AND NOT (#MainStep.S57)) AND ("DB720_KuKa_MainCtrl".CmdOut.gi_ToolTypeNo <> 2))) AND "DB1900_Communication_PC".Para.DiamondVibCylinder) AND NOT ("DB1080_Component".Robot.Status.Busy) 成立时，将 TRUE 传送到 #DiamondAutoStep.DiamondStep.StartCmd
   IF ((((#MainStep.S44 AND NOT (#MainStep.S57)) AND ("DB720_KuKa_MainCtrl".CmdOut.gi_ToolTypeNo <> 2))) AND "DB1900_Communication_PC".Para.DiamondVibCylinder) AND NOT ("DB1080_Component".Robot.Status.Busy) THEN
       #DiamondAutoStep.DiamondStep.StartCmd := TRUE;
   END_IF;
   // 含义：将 (#MainStep.S44 AND #DiamondAutoStep.DiamondStep.StartCmd) OR (#MainStep.S44 AND #MainStep.S57) 赋给 #MainStep.S57
   #MainStep.S57 := (#MainStep.S44 AND #DiamondAutoStep.DiamondStep.StartCmd) OR (#MainStep.S44 AND #MainStep.S57);
   // 含义：将 ((#MainStep.S44 AND ("DB720_KuKa_MainCtrl".CmdOut.gi_ToolTypeNo = 2))) OR (((#MainStep.S44 AND ("DB720_KuKa_MainCtrl".CmdOut.gi_ToolTypeNo <> 2))) AND NOT ("DB1900_Communication_PC".Para.DiamondVibCylinder)) 赋给 #MainStep.S58
   #MainStep.S58 := ((#MainStep.S44 AND ("DB720_KuKa_MainCtrl".CmdOut.gi_ToolTypeNo = 2))) OR (((#MainStep.S44 AND ("DB720_KuKa_MainCtrl".CmdOut.gi_ToolTypeNo <> 2))) AND NOT ("DB1900_Communication_PC".Para.DiamondVibCylinder));

   // ---------- 网络 28 ----------
   // 含义：将 (#MainStep.S57 AND #DiamondAutoStep.DiamondStep.TaskIO) OR (#MainStep.S57 AND #DiamondAutoStep.DiamondStep.TaskIO) OR (#MainStep.S57 AND #MainStep.S59) 赋给 #MainStep.S59
   #MainStep.S59 := (#MainStep.S57 AND #DiamondAutoStep.DiamondStep.TaskIO) OR (#MainStep.S57 AND #DiamondAutoStep.DiamondStep.TaskIO) OR (#MainStep.S57 AND #MainStep.S59);

   // ---------- 网络 29 ----------
   // 标题：放工具冷却
   // 含义：条件 (((((#MainStep.S44 OR #MainStep.S58 OR #MainStep.S59) AND NOT (#MainStep.S45)) AND "DB1080_Component".Robot.Status.HomePos) AND "DB1900_Communication_PC".Recv.WorkStart) AND ("DB720_KuKa_MainCtrl".CmdOut.gi_ToolTypeNo = 2)) 成立时，将 TRUE 传送到 #RobotAutoStep.Cmd.Auto.ChangeTool
   IF (((((#MainStep.S44 OR #MainStep.S58 OR #MainStep.S59) AND NOT (#MainStep.S45)) AND "DB1080_Component".Robot.Status.HomePos) AND "DB1900_Communication_PC".Recv.WorkStart) AND ("DB720_KuKa_MainCtrl".CmdOut.gi_ToolTypeNo = 2)) THEN
       #RobotAutoStep.Cmd.Auto.ChangeTool := TRUE;
   END_IF;
   // 含义：条件 ((((((#MainStep.S44 OR #MainStep.S58 OR #MainStep.S59) AND NOT (#MainStep.S45)) AND "DB1080_Component".Robot.Status.HomePos) AND "DB1900_Communication_PC".Recv.WorkStart) AND ("DB720_KuKa_MainCtrl".CmdOut.gi_ToolTypeNo <> 2))) AND "DB1900_Communication_PC".Para.DiamondVibCylinder 成立时，将 TRUE 传送到 #DiamondAutoStep.DiamondStep.StartCmd
   IF ((((((#MainStep.S44 OR #MainStep.S58 OR #MainStep.S59) AND NOT (#MainStep.S45)) AND "DB1080_Component".Robot.Status.HomePos) AND "DB1900_Communication_PC".Recv.WorkStart) AND ("DB720_KuKa_MainCtrl".CmdOut.gi_ToolTypeNo <> 2))) AND "DB1900_Communication_PC".Para.DiamondVibCylinder THEN
       #DiamondAutoStep.DiamondStep.StartCmd := TRUE;
   END_IF;
   // 含义：将 (((((#MainStep.S44 OR #MainStep.S58 OR #MainStep.S59) AND ("DB720_KuKa_MainCtrl".CmdOut.gi_ToolTypeNo = 2))) AND #RobotAutoStep.ChangeToolStatus.TaskDone) AND #RobotAutoStep.ChangeToolStatus.TaskIO) OR ((((((#MainStep.S44 OR #MainStep.S58 OR #MainStep.S59) AND ("DB720_KuKa_MainCtrl".CmdOut.gi_ToolTypeNo <> 2))) AND "DB1900_Communication_PC".Para.DiamondVibCylinder) AND #DiamondAutoStep.DiamondStep.TaskDone) AND #DiamondAutoStep.DiamondStep.TaskIO) OR ((((#MainStep.S44 OR #MainStep.S58 OR #MainStep.S59) AND ("DB720_KuKa_MainCtrl".CmdOut.gi_ToolTypeNo <> 2))) AND NOT ("DB1900_Communication_PC".Para.DiamondVibCylinder)) OR ((#MainStep.S44 OR #MainStep.S58 OR #MainStep.S59) AND #MainStep.S45) 赋给 #MainStep.S45
   #MainStep.S45 := (((((#MainStep.S44 OR #MainStep.S58 OR #MainStep.S59) AND ("DB720_KuKa_MainCtrl".CmdOut.gi_ToolTypeNo = 2))) AND #RobotAutoStep.ChangeToolStatus.TaskDone) AND #RobotAutoStep.ChangeToolStatus.TaskIO) OR ((((((#MainStep.S44 OR #MainStep.S58 OR #MainStep.S59) AND ("DB720_KuKa_MainCtrl".CmdOut.gi_ToolTypeNo <> 2))) AND "DB1900_Communication_PC".Para.DiamondVibCylinder) AND #DiamondAutoStep.DiamondStep.TaskDone) AND #DiamondAutoStep.DiamondStep.TaskIO) OR ((((#MainStep.S44 OR #MainStep.S58 OR #MainStep.S59) AND ("DB720_KuKa_MainCtrl".CmdOut.gi_ToolTypeNo <> 2))) AND NOT ("DB1900_Communication_PC".Para.DiamondVibCylinder)) OR ((#MainStep.S44 OR #MainStep.S58 OR #MainStep.S59) AND #MainStep.S45);

   // ---------- 网络 30 ----------
   // 标题：换枪
   // 含义：条件 (((#MainStep.S45 AND NOT (#MainStep.S46)) AND "DB720_KuKa_MainCtrl".Aux.ToolAtPosTimer.Q) AND ("DB720_KuKa_MainCtrl".CmdOut.gi_ToolTypeNo = 2)) 成立时，将 TRUE 传送到 "DB1080_Component".Robot.Cmd.Auto.GoHome
   IF (((#MainStep.S45 AND NOT (#MainStep.S46)) AND "DB720_KuKa_MainCtrl".Aux.ToolAtPosTimer.Q) AND ("DB720_KuKa_MainCtrl".CmdOut.gi_ToolTypeNo = 2)) THEN
       "DB1080_Component".Robot.Cmd.Auto.GoHome := TRUE;
   END_IF;
   // 含义：将 (((#MainStep.S45 AND "DB1080_Component".Robot.Status.HomePos) OR (#MainStep.S45 AND NOT ("DB720_KuKa_MainCtrl".Aux.ToolAtPosTimer.Q)) OR ((#MainStep.S45 AND ("DB720_KuKa_MainCtrl".CmdOut.gi_ToolTypeNo <> 2))) OR (#MainStep.S45 AND #MainStep.S46)) AND "DB1900_Communication_PC".Recv.ChangeTool) OR ((((#MainStep.S45 AND "DB1080_Component".Robot.Status.HomePos) OR (#MainStep.S45 AND NOT ("DB720_KuKa_MainCtrl".Aux.ToolAtPosTimer.Q)) OR ((#MainStep.S45 AND ("DB720_KuKa_MainCtrl".CmdOut.gi_ToolTypeNo <> 2))) OR (#MainStep.S45 AND #MainStep.S46)) AND ("DB720_KuKa_MainCtrl".CmdOut.gi_ToolTypeNo <> 2))) 赋给 #MainStep.S46
   #MainStep.S46 := (((#MainStep.S45 AND "DB1080_Component".Robot.Status.HomePos) OR (#MainStep.S45 AND NOT ("DB720_KuKa_MainCtrl".Aux.ToolAtPosTimer.Q)) OR ((#MainStep.S45 AND ("DB720_KuKa_MainCtrl".CmdOut.gi_ToolTypeNo <> 2))) OR (#MainStep.S45 AND #MainStep.S46)) AND "DB1900_Communication_PC".Recv.ChangeTool) OR ((((#MainStep.S45 AND "DB1080_Component".Robot.Status.HomePos) OR (#MainStep.S45 AND NOT ("DB720_KuKa_MainCtrl".Aux.ToolAtPosTimer.Q)) OR ((#MainStep.S45 AND ("DB720_KuKa_MainCtrl".CmdOut.gi_ToolTypeNo <> 2))) OR (#MainStep.S45 AND #MainStep.S46)) AND ("DB720_KuKa_MainCtrl".CmdOut.gi_ToolTypeNo <> 2)));
   // 含义：条件 (#MainStep.S45 AND "DB1080_Component".Robot.Status.HomePos) OR (#MainStep.S45 AND NOT ("DB720_KuKa_MainCtrl".Aux.ToolAtPosTimer.Q)) OR ((#MainStep.S45 AND ("DB720_KuKa_MainCtrl".CmdOut.gi_ToolTypeNo <> 2))) OR (#MainStep.S45 AND #MainStep.S46) 成立时，将 0.5 传送到 "DB1080_Component".Aux.Pressure
   IF (#MainStep.S45 AND "DB1080_Component".Robot.Status.HomePos) OR (#MainStep.S45 AND NOT ("DB720_KuKa_MainCtrl".Aux.ToolAtPosTimer.Q)) OR ((#MainStep.S45 AND ("DB720_KuKa_MainCtrl".CmdOut.gi_ToolTypeNo <> 2))) OR (#MainStep.S45 AND #MainStep.S46) THEN
       "DB1080_Component".Aux.Pressure := 0.5;
   END_IF;

   // ---------- 网络 31 ----------
   // 含义：将 (#MainStep.S46 AND NOT ("DB1080_Component".Robot.Status.Busy)) OR (#MainStep.S46 AND #MainStep.S47) 赋给 #MainStep.S47
   #MainStep.S47 := (#MainStep.S46 AND NOT ("DB1080_Component".Robot.Status.Busy)) OR (#MainStep.S46 AND #MainStep.S47);
   // 含义：条件 #MainStep.S46 AND NOT (#MainStep.S47) 成立时，将 FALSE 传送到 #RobotAutoStep.ChangeToolStatus.TaskDone
   IF #MainStep.S46 AND NOT (#MainStep.S47) THEN
       #RobotAutoStep.ChangeToolStatus.TaskDone := FALSE;
   END_IF;

   // ---------- 网络 32 ----------
   // 标题：请求上位机参数录入...
   // 含义：条件 #MainStep.S47 AND NOT (#MainStep.S48) 成立时，将 TRUE 传送到 "DB1081_ValveCall".ST01.Z08.ExtAuto
   IF #MainStep.S47 AND NOT (#MainStep.S48) THEN
       "DB1081_ValveCall".ST01.Z08.ExtAuto := TRUE;
   END_IF;
   // 含义：将 ((#MainStep.S47 AND "DB1900_Communication_PC".Recv.ParaWriteDone) AND "DB1081_ValveCall".ST01.Z08.ExtPos) OR (#MainStep.S47 AND #MainStep.S48) 赋给 #MainStep.S48
   #MainStep.S48 := ((#MainStep.S47 AND "DB1900_Communication_PC".Recv.ParaWriteDone) AND "DB1081_ValveCall".ST01.Z08.ExtPos) OR (#MainStep.S47 AND #MainStep.S48);

   // ---------- 网络 33 ----------
   // 标题：检查是否需要换型
   // 含义：将 ((#MainStep.S48 AND ("DB1900_Communication_PC".Para.IOFixtureNo <> "DB1080_Component".IOFixtureIID.TP_CurFixtureID))) OR ((#MainStep.S48 AND ("DB1900_Communication_PC".Para.PowerFixtureNo <> "DB1080_Component".PowerFixtureID.TP_CurFixtureID))) OR (#MainStep.S48 AND #MainStep.S49) 赋给 #MainStep.S49
   #MainStep.S49 := ((#MainStep.S48 AND ("DB1900_Communication_PC".Para.IOFixtureNo <> "DB1080_Component".IOFixtureIID.TP_CurFixtureID))) OR ((#MainStep.S48 AND ("DB1900_Communication_PC".Para.PowerFixtureNo <> "DB1080_Component".PowerFixtureID.TP_CurFixtureID))) OR (#MainStep.S48 AND #MainStep.S49);
   // 含义：将 (((((#MainStep.S48 AND NOT (#MainStep.S49)) AND ("DB1900_Communication_PC".Para.IOFixtureNo = "DB1080_Component".IOFixtureIID.TP_CurFixtureID))) AND ("DB1900_Communication_PC".Para.PowerFixtureNo = "DB1080_Component".PowerFixtureID.TP_CurFixtureID))) OR (#MainStep.S48 AND #EdgeDetc.Pulse[0]) 赋给 #EdgeDetc.Pulse[0]
   #EdgeDetc.Pulse[0] := (((((#MainStep.S48 AND NOT (#MainStep.S49)) AND ("DB1900_Communication_PC".Para.IOFixtureNo = "DB1080_Component".IOFixtureIID.TP_CurFixtureID))) AND ("DB1900_Communication_PC".Para.PowerFixtureNo = "DB1080_Component".PowerFixtureID.TP_CurFixtureID))) OR (#MainStep.S48 AND #EdgeDetc.Pulse[0]);

   // ---------- 网络 34 ----------
   // 标题：换枪
   // 含义：条件 ((#MainStep.S49 AND NOT (#EdgeDetc.Pulse[0])) AND ("DB720_KuKa_MainCtrl".CmdOut.gi_ToolTypeNo = 2)) 成立时，将 TRUE 传送到 #RobotAutoStep.Cmd.Auto.ChangeTool
   IF ((#MainStep.S49 AND NOT (#EdgeDetc.Pulse[0])) AND ("DB720_KuKa_MainCtrl".CmdOut.gi_ToolTypeNo = 2)) THEN
       #RobotAutoStep.Cmd.Auto.ChangeTool := TRUE;
   END_IF;
   // 含义：将 ((#MainStep.S49 AND #RobotAutoStep.ChangeToolStatus.TaskDone) AND #RobotAutoStep.ChangeToolStatus.TaskIO) OR (#MainStep.S49 AND #EdgeDetc.Pulse[0]) 赋给 #EdgeDetc.Pulse[0]
   #EdgeDetc.Pulse[0] := ((#MainStep.S49 AND #RobotAutoStep.ChangeToolStatus.TaskDone) AND #RobotAutoStep.ChangeToolStatus.TaskIO) OR (#MainStep.S49 AND #EdgeDetc.Pulse[0]);

   // ---------- 网络 35 ----------
   // 含义：将 (#MainStep.S50 AND NOT ("DB1080_Component".Robot.Status.Busy)) OR (#MainStep.S50 AND #MainStep.S51) 赋给 #MainStep.S51
   #MainStep.S51 := (#MainStep.S50 AND NOT ("DB1080_Component".Robot.Status.Busy)) OR (#MainStep.S50 AND #MainStep.S51);

   // ---------- 网络 36 ----------
   // 含义：条件 #MainStep.S51 AND NOT (#MainStep.S52) 成立时，将 TRUE 传送到 "DB1080_Component".Robot.Cmd.Auto.GoHome
   IF #MainStep.S51 AND NOT (#MainStep.S52) THEN
       "DB1080_Component".Robot.Cmd.Auto.GoHome := TRUE;
   END_IF;
   // 含义：将 (#MainStep.S51 AND "DB1080_Component".Robot.Status.HomePos) OR (#MainStep.S51 AND #MainStep.S52) 赋给 #MainStep.S52
   #MainStep.S52 := (#MainStep.S51 AND "DB1080_Component".Robot.Status.HomePos) OR (#MainStep.S51 AND #MainStep.S52);
   // 含义：条件 (#MainStep.S51 AND "DB1080_Component".Robot.Status.HomePos) OR (#MainStep.S51 AND #MainStep.S52) 成立时，将 0.5 传送到 "DB1080_Component".Aux.Pressure
   IF (#MainStep.S51 AND "DB1080_Component".Robot.Status.HomePos) OR (#MainStep.S51 AND #MainStep.S52) THEN
       "DB1080_Component".Aux.Pressure := 0.5;
   END_IF;

   // ---------- 网络 37 ----------
   // 标题：换枪
   // 含义：条件 ((#MainStep.S52 AND "DB1080_Component".Robot.Status.HomePos) AND ("DB720_KuKa_MainCtrl".CmdOut.gi_ToolTypeNo = 2)) 成立时，将 TRUE 传送到 #RobotAutoStep.Cmd.Auto.ChangeTool
   IF ((#MainStep.S52 AND "DB1080_Component".Robot.Status.HomePos) AND ("DB720_KuKa_MainCtrl".CmdOut.gi_ToolTypeNo = 2)) THEN
       #RobotAutoStep.Cmd.Auto.ChangeTool := TRUE;
   END_IF;
   // 含义：将 (#MainStep.S52 AND "DB1080_Component".Robot.Status.HomePos) AND "DB1900_Communication_PC".Recv.WorkDone 赋给 "DB1900_Communication_PC".Send.WorkDone
   "DB1900_Communication_PC".Send.WorkDone := (#MainStep.S52 AND "DB1080_Component".Robot.Status.HomePos) AND "DB1900_Communication_PC".Recv.WorkDone;
   // 含义：将 (#MainStep.S52 AND #RobotAutoStep.ChangeToolStatus.TaskDone) AND #RobotAutoStep.ChangeToolStatus.TaskIO 赋给 #MainStep.S53
   #MainStep.S53 := (#MainStep.S52 AND #RobotAutoStep.ChangeToolStatus.TaskDone) AND #RobotAutoStep.ChangeToolStatus.TaskIO;

   // ---------- 网络 38 ----------
   // 标题：自动步结束
   // 含义：将 #MainStep.S53 OR #MainStep.ErrEnd 赋给 #MainStep.End
   #MainStep.End := #MainStep.S53 OR #MainStep.ErrEnd;
   // 含义：条件 #MainStep.S53 OR #MainStep.ErrEnd 成立时，将 0.5 传送到 "DB1080_Component".Aux.Pressure
   IF #MainStep.S53 OR #MainStep.ErrEnd THEN
       "DB1080_Component".Aux.Pressure := 0.5;
   END_IF;

   // ---------- 网络 39 ----------
   // 含义：调用块/实例 #RobotAutoStep
   #RobotAutoStep();

   // ---------- 网络 40 ----------
   // 标题：HorDrillAutoStep
   // 含义：调用块/实例 #HorDrillAutoStep
   #HorDrillAutoStep();

   // ---------- 网络 41 ----------
   // 标题：DownDrillAutoStep
   // 含义：调用块/实例 #DownDrillAutoStep
   #DownDrillAutoStep();

   // ---------- 网络 42 ----------
   // 标题：CoreDrillAutoStep
   // 含义：调用块/实例 #DiamondAutoStep
   #DiamondAutoStep();

   // ---------- 网络 43 ----------
   // （空白网络）
END_FUNCTION_BLOCK

FUNCTION_BLOCK "FB1061_RobotAutoStep"   // FB1061, SCL
{ S7_Optimized_Access := 'TRUE' }
// ============================================================
//  Block: FB1061_RobotAutoStep
//  ============================================================
//  编号：FB1061
//  原始语言：LAD（规则翻译为 SCL）
//  含义：自动循环起点
   VAR_INPUT
      StepStart : Bool;   // 输入参数
   END_VAR
   VAR
      Cmd : Struct   // 静态变量
         Auto : Struct   // 静态变量
            Drill : Bool;   // 钻孔
            CheckBit : Bool;   // 校验
            ChangeTool : Bool;   // 换枪
         END_STRUCT;
      END_STRUCT;
      AtCmd : Word;   // 静态变量
      Status : Struct   // 静态变量
         Running : Bool;   // 自动运行中
         OkToStart : Bool;   // 设备可以启动
         OKPartPrompt : Bool;   // 结果OK
         NGPartPrompt : Bool;   // 结果NG
         ToBeHomePos : Bool;   // 回原点提示
         AllStationDone : Bool;   // 所有工位完成
         SP6 : Bool;   // 静态变量
         SP7 : Bool;   // 静态变量
         SP : Byte;   // 静态变量
      END_STRUCT;
      AtStatus : Word;   // 静态变量
      DrillStatus : Struct   // 静态变量
         OkToStart : Bool;   // 静态变量
         Busy : Bool;   // 静态变量
         TaskDone : Bool;   // 静态变量
         TaskIO : Bool;   // 静态变量
         TaskNIO : Bool;   // 静态变量
      END_STRUCT;
      ATDrillStatus : Word;   // 静态变量
      CheckBitStatus : Struct   // 静态变量
         OkToStart : Bool;   // 静态变量
         Busy : Bool;   // 静态变量
         TaskDone : Bool;   // 静态变量
         TaskIO : Bool;   // 静态变量
         TaskNIO : Bool;   // 静态变量
      END_STRUCT;
      AT : Word;   // 静态变量
      ChangeToolStatus : Struct   // 静态变量
         OkToStart : Bool;   // 静态变量
         Busy : Bool;   // 静态变量
         TaskDone : Bool;   // 静态变量
         TaskIO : Bool;   // 静态变量
         TaskNIO : Bool;   // 静态变量
      END_STRUCT;
      AtChangeToolStatus : Word;   // 静态变量
      EdgeDetc : Struct   // 静态变量
         Pulse : Array[0..15] of Bool;   // 静态变量
      END_STRUCT;
      MainStep : "UDT_Step";   // 自动流程步
      CycleTime : "FB5008_CycleTime";   // 静态变量
      StartCmd_ManMode : Bool;   // 静态变量
      StartCmd_AutoMode : Bool;   // 静态变量
      OkToStart : Bool;   // 静态变量
      HomePos : Bool;   // 静态变量
      "Do" : Bool;   // 静态变量
      Done : Bool;   // 静态变量
      PartOn : Bool;   // 静态变量
      PartOK : Bool;   // 静态变量
      PartNG : Bool;   // 静态变量
      Start : Bool;   // 静态变量
      End : Bool;   // 静态变量
      ErrEnd : Bool;   // 静态变量
      S1 : Bool;   // 静态变量
      S2 : Bool;   // 静态变量
      S3 : Bool;   // 静态变量
      S4 : Bool;   // 静态变量
      S5 : Bool;   // 静态变量
      S6 : Bool;   // 静态变量
      S7 : Bool;   // 静态变量
      S8 : Bool;   // 静态变量
      S9 : Bool;   // 静态变量
      S10 : Bool;   // 静态变量
      S11 : Bool;   // 静态变量
      S12 : Bool;   // 静态变量
      S13 : Bool;   // 静态变量
      S14 : Bool;   // 静态变量
      S15 : Bool;   // 静态变量
      S16 : Bool;   // 静态变量
      S17 : Bool;   // 静态变量
      S18 : Bool;   // 静态变量
      S19 : Bool;   // 静态变量
      S20 : Bool;   // 静态变量
      S21 : Bool;   // 静态变量
      S22 : Bool;   // 静态变量
      S23 : Bool;   // 静态变量
      S24 : Bool;   // 静态变量
      S25 : Bool;   // 静态变量
      S26 : Bool;   // 静态变量
      S27 : Bool;   // 静态变量
      S28 : Bool;   // 静态变量
      S29 : Bool;   // 静态变量
      S30 : Bool;   // 静态变量
      S31 : Bool;   // 静态变量
      S32 : Bool;   // 静态变量
      S33 : Bool;   // 静态变量
      S34 : Bool;   // 静态变量
      S35 : Bool;   // 静态变量
      S36 : Bool;   // 静态变量
      S37 : Bool;   // 静态变量
      S38 : Bool;   // 静态变量
      S39 : Bool;   // 静态变量
      S40 : Bool;   // 静态变量
      S41 : Bool;   // 静态变量
      S42 : Bool;   // 静态变量
      S43 : Bool;   // 静态变量
      S44 : Bool;   // 静态变量
      S45 : Bool;   // 静态变量
      S46 : Bool;   // 静态变量
      S47 : Bool;   // 静态变量
      S48 : Bool;   // 静态变量
      S49 : Bool;   // 静态变量
      S50 : Bool;   // 静态变量
      S51 : Bool;   // 静态变量
      S52 : Bool;   // 静态变量
      S53 : Bool;   // 静态变量
      S54 : Bool;   // 静态变量
      S55 : Bool;   // 静态变量
      S56 : Bool;   // 静态变量
      S57 : Bool;   // 静态变量
      S58 : Bool;   // 静态变量
      S59 : Bool;   // 静态变量
      S60 : Bool;   // 静态变量
      S61 : Bool;   // 静态变量
      S62 : Bool;   // 静态变量
      S63 : Bool;   // 静态变量
      S64 : Bool;   // 静态变量
      S65 : Bool;   // 静态变量
      S66 : Bool;   // 静态变量
      S67 : Bool;   // 静态变量
      CycleTime_Net : Time;   // 静态变量
      CycleTime_Total : Time;   // 静态变量
      Aux : Struct   // 静态变量
         StartPls : Bool;   // 静态变量
         EndPls : Bool;   // 静态变量
         sp : Byte;   // 静态变量
         StartTime : Time_Of_Day;   // 静态变量
         LastEndTime : Time_Of_Day;   // 静态变量
      END_STRUCT;
   END_VAR
   VAR_TEMP
      StepPls : Bool;   // 临时变量
   END_VAR
BEGIN

   // ---------- 网络 1 ----------
   // 标题：模式分配
   // 含义：将 ("StepMode_M" AND "DB1001_SysMode".SubSysMode.Mode.StepPls) OR ("StepMode_M" AND #MainStep.StartCmd_ManMode) OR "ManMode_M" OR "AutoMode_M" 赋给 #StepPls
   #StepPls := ("StepMode_M" AND "DB1001_SysMode".SubSysMode.Mode.StepPls) OR ("StepMode_M" AND #MainStep.StartCmd_ManMode) OR "ManMode_M" OR "AutoMode_M";

   // ---------- 网络 2 ----------
   // 标题：提示回原点
   // 含义：将 "ASMMode_M" AND NOT ("DB1001_SysMode".SubSysMode.Status.ErrPresent) 赋给 #Status.OkToStart
   #Status.OkToStart := "ASMMode_M" AND NOT ("DB1001_SysMode".SubSysMode.Status.ErrPresent);
   // 含义：将 #DrillStatus.Busy OR #ChangeToolStatus.Busy OR #CheckBitStatus.Busy 赋给 #Status.Running
   #Status.Running := #DrillStatus.Busy OR #ChangeToolStatus.Busy OR #CheckBitStatus.Busy;

   // ---------- 网络 3 ----------
   // 标题：自动步开始
   // 注释：自动循环起点
   // 含义：将 ((((#Status.OkToStart OR #MainStep.Start) AND "ASMMode_M") AND NOT ("DB1900_Communication_PC".Recv.EmmMode)) AND NOT ("DB1040_HomePos".MainStep.Start)) AND NOT (#MainStep.End) 赋给 #MainStep.Start
   #MainStep.Start := ((((#Status.OkToStart OR #MainStep.Start) AND "ASMMode_M") AND NOT ("DB1900_Communication_PC".Recv.EmmMode)) AND NOT ("DB1040_HomePos".MainStep.Start)) AND NOT (#MainStep.End);
   // 含义：条件 NOT (#Status.OkToStart OR #MainStep.Start) 成立时，将 FALSE 传送到 #MainStep.ErrEnd
   IF NOT (#Status.OkToStart OR #MainStep.Start) THEN
       #MainStep.ErrEnd := FALSE;
   END_IF;
   // 含义：条件 NOT (#Status.OkToStart OR #MainStep.Start) 成立时，将 FALSE 传送到 #DrillStatus.Busy
   IF NOT (#Status.OkToStart OR #MainStep.Start) THEN
       #DrillStatus.Busy := FALSE;
   END_IF;
   // 含义：条件 NOT (#Status.OkToStart OR #MainStep.Start) 成立时，将 FALSE 传送到 #ChangeToolStatus.Busy
   IF NOT (#Status.OkToStart OR #MainStep.Start) THEN
       #ChangeToolStatus.Busy := FALSE;
   END_IF;
   // 含义：条件 NOT (#Status.OkToStart OR #MainStep.Start) 成立时，将 FALSE 传送到 #CheckBitStatus.Busy
   IF NOT (#Status.OkToStart OR #MainStep.Start) THEN
       #CheckBitStatus.Busy := FALSE;
   END_IF;
   // 含义：条件 NOT (#Status.OkToStart OR #MainStep.Start) 成立时，将 FALSE 传送到 #CheckBitStatus.TaskDone
   IF NOT (#Status.OkToStart OR #MainStep.Start) THEN
       #CheckBitStatus.TaskDone := FALSE;
   END_IF;
   // 含义：条件 NOT (#Status.OkToStart OR #MainStep.Start) 成立时，将 FALSE 传送到 #ChangeToolStatus.TaskDone
   IF NOT (#Status.OkToStart OR #MainStep.Start) THEN
       #ChangeToolStatus.TaskDone := FALSE;
   END_IF;
   // 含义：条件 NOT (#Status.OkToStart OR #MainStep.Start) 成立时，将 FALSE 传送到 #DrillStatus.TaskDone
   IF NOT (#Status.OkToStart OR #MainStep.Start) THEN
       #DrillStatus.TaskDone := FALSE;
   END_IF;

   // ---------- 网络 4 ----------
   // 标题：有故障，断开正常流程，转入故障处理；
   // 含义：条件 #MainStep.Start AND NOT (#MainStep.S1) 成立时，将 0 传送到 #ATDrillStatus
   IF #MainStep.Start AND NOT (#MainStep.S1) THEN
       #ATDrillStatus := 0;
   END_IF;
   // 含义：条件 #MainStep.Start AND NOT (#MainStep.S1) 成立时，将 FALSE 传送到 #DrillStatus.Busy
   IF #MainStep.Start AND NOT (#MainStep.S1) THEN
       #DrillStatus.Busy := FALSE;
   END_IF;
   // 含义：将 #MainStep.Start AND NOT (#MainStep.ErrEnd) 赋给 #MainStep.S1
   #MainStep.S1 := #MainStep.Start AND NOT (#MainStep.ErrEnd);

   // ---------- 网络 5 ----------
   // 含义：当 #MainStep.S1 为 TRUE 时置位 #MainStep.S2，否则复位（触点→线圈）
   IF #MainStep.S1 THEN
       #MainStep.S2 := TRUE;
   ELSE
       #MainStep.S2 := FALSE;
   END_IF;

   // ---------- 网络 6 ----------
   // 标题：流程分支
   // 含义：将 ((((((#MainStep.S2 AND #Cmd.Auto.ChangeTool) AND NOT ("DB1080_Component".Robot.Status.Busy)) OR (#MainStep.S2 AND #EdgeDetc.Pulse[0])) AND NOT (#EdgeDetc.Pulse[0])) AND NOT (#EdgeDetc.Pulse[0])) AND NOT (#EdgeDetc.Pulse[0])) AND NOT (#EdgeDetc.Pulse[0]) 赋给 #EdgeDetc.Pulse[0]
   #EdgeDetc.Pulse[0] := ((((((#MainStep.S2 AND #Cmd.Auto.ChangeTool) AND NOT ("DB1080_Component".Robot.Status.Busy)) OR (#MainStep.S2 AND #EdgeDetc.Pulse[0])) AND NOT (#EdgeDetc.Pulse[0])) AND NOT (#EdgeDetc.Pulse[0])) AND NOT (#EdgeDetc.Pulse[0])) AND NOT (#EdgeDetc.Pulse[0]);
   // 含义：将 (((((((#MainStep.S2 AND #Cmd.Auto.Drill) AND NOT ("DB1080_Component".Robot.Status.Busy)) AND "DB1900_Communication_PC".Para.DrillDirection1) OR (#MainStep.S2 AND #EdgeDetc.Pulse[0])) AND NOT (#EdgeDetc.Pulse[0])) AND NOT (#EdgeDetc.Pulse[0])) AND NOT (#EdgeDetc.Pulse[0])) AND NOT (#EdgeDetc.Pulse[0]) 赋给 #EdgeDetc.Pulse[0]
   #EdgeDetc.Pulse[0] := (((((((#MainStep.S2 AND #Cmd.Auto.Drill) AND NOT ("DB1080_Component".Robot.Status.Busy)) AND "DB1900_Communication_PC".Para.DrillDirection1) OR (#MainStep.S2 AND #EdgeDetc.Pulse[0])) AND NOT (#EdgeDetc.Pulse[0])) AND NOT (#EdgeDetc.Pulse[0])) AND NOT (#EdgeDetc.Pulse[0])) AND NOT (#EdgeDetc.Pulse[0]);
   // 含义：将 (((((((#MainStep.S2 AND #Cmd.Auto.Drill) AND NOT ("DB1080_Component".Robot.Status.Busy)) AND "DB1900_Communication_PC".Para.DrillDirection3) OR (#MainStep.S2 AND #EdgeDetc.Pulse[0])) AND NOT (#EdgeDetc.Pulse[0])) AND NOT (#EdgeDetc.Pulse[0])) AND NOT (#EdgeDetc.Pulse[0])) AND NOT (#EdgeDetc.Pulse[0]) 赋给 #EdgeDetc.Pulse[0]
   #EdgeDetc.Pulse[0] := (((((((#MainStep.S2 AND #Cmd.Auto.Drill) AND NOT ("DB1080_Component".Robot.Status.Busy)) AND "DB1900_Communication_PC".Para.DrillDirection3) OR (#MainStep.S2 AND #EdgeDetc.Pulse[0])) AND NOT (#EdgeDetc.Pulse[0])) AND NOT (#EdgeDetc.Pulse[0])) AND NOT (#EdgeDetc.Pulse[0])) AND NOT (#EdgeDetc.Pulse[0]);
   // 含义：将 ((((((#MainStep.S2 AND #Cmd.Auto.CheckBit) AND NOT ("DB1080_Component".Robot.Status.Busy)) OR (#MainStep.S2 AND #EdgeDetc.Pulse[0])) AND NOT (#EdgeDetc.Pulse[0])) AND NOT (#EdgeDetc.Pulse[0])) AND NOT (#EdgeDetc.Pulse[0])) AND NOT (#EdgeDetc.Pulse[0]) 赋给 #EdgeDetc.Pulse[0]
   #EdgeDetc.Pulse[0] := ((((((#MainStep.S2 AND #Cmd.Auto.CheckBit) AND NOT ("DB1080_Component".Robot.Status.Busy)) OR (#MainStep.S2 AND #EdgeDetc.Pulse[0])) AND NOT (#EdgeDetc.Pulse[0])) AND NOT (#EdgeDetc.Pulse[0])) AND NOT (#EdgeDetc.Pulse[0])) AND NOT (#EdgeDetc.Pulse[0]);

   // ---------- 网络 7 ----------
   // 标题：查看机器人状态
   // 含义：条件 #EdgeDetc.Pulse[0] AND NOT (#MainStep.S3) 成立时，将 TRUE 传送到 #ChangeToolStatus.Busy
   IF #EdgeDetc.Pulse[0] AND NOT (#MainStep.S3) THEN
       #ChangeToolStatus.Busy := TRUE;
   END_IF;
   // 含义：条件 #EdgeDetc.Pulse[0] AND NOT (#MainStep.S3) 成立时，将 FALSE 传送到 #ChangeToolStatus.TaskIO
   IF #EdgeDetc.Pulse[0] AND NOT (#MainStep.S3) THEN
       #ChangeToolStatus.TaskIO := FALSE;
   END_IF;
   // 含义：将 (#EdgeDetc.Pulse[0] AND NOT ("DB720_KuKa_MainCtrl".ChangeTool.Busy)) OR (#EdgeDetc.Pulse[0] AND #MainStep.S7) 赋给 #MainStep.S7
   #MainStep.S7 := (#EdgeDetc.Pulse[0] AND NOT ("DB720_KuKa_MainCtrl".ChangeTool.Busy)) OR (#EdgeDetc.Pulse[0] AND #MainStep.S7);

   // ---------- 网络 8 ----------
   // 标题：****************************开始换夹具*******************************
   // 含义：条件 #MainStep.S7 AND NOT (#MainStep.S9) 成立时，将 TRUE 传送到 "DB720_KuKa_MainCtrl".ChangeTool.StartCmd
   IF #MainStep.S7 AND NOT (#MainStep.S9) THEN
       "DB720_KuKa_MainCtrl".ChangeTool.StartCmd := TRUE;
   END_IF;
   // 含义：将 ((#MainStep.S7 AND "DB720_KuKa_MainCtrl".ChangeTool.TaskDone) AND "DB720_KuKa_MainCtrl".ChangeTool.TaskIO) OR (#MainStep.S7 AND #MainStep.S9) 赋给 #MainStep.S9
   #MainStep.S9 := ((#MainStep.S7 AND "DB720_KuKa_MainCtrl".ChangeTool.TaskDone) AND "DB720_KuKa_MainCtrl".ChangeTool.TaskIO) OR (#MainStep.S7 AND #MainStep.S9);

   // ---------- 网络 9 ----------
   // 标题：换夹具结束
   // 含义：条件 #MainStep.S9 AND NOT (#MainStep.S11) 成立时，将 TRUE 传送到 #ChangeToolStatus.TaskDone
   IF #MainStep.S9 AND NOT (#MainStep.S11) THEN
       #ChangeToolStatus.TaskDone := TRUE;
   END_IF;
   // 含义：条件 #MainStep.S9 AND NOT (#MainStep.S11) 成立时，将 TRUE 传送到 #ChangeToolStatus.TaskIO
   IF #MainStep.S9 AND NOT (#MainStep.S11) THEN
       #ChangeToolStatus.TaskIO := TRUE;
   END_IF;
   // 含义：将 (#MainStep.S9 AND NOT (#Cmd.Auto.ChangeTool)) OR (#MainStep.S9 AND #MainStep.S11) 赋给 #MainStep.S11
   #MainStep.S11 := (#MainStep.S9 AND NOT (#Cmd.Auto.ChangeTool)) OR (#MainStep.S9 AND #MainStep.S11);

   // ---------- 网络 10 ----------
   // 标题：检查机器人状态
   // 含义：条件 #EdgeDetc.Pulse[0] AND NOT (#MainStep.S15) 成立时，将 TRUE 传送到 #DrillStatus.Busy
   IF #EdgeDetc.Pulse[0] AND NOT (#MainStep.S15) THEN
       #DrillStatus.Busy := TRUE;
   END_IF;
   // 含义：条件 #EdgeDetc.Pulse[0] AND NOT (#MainStep.S15) 成立时，将 FALSE 传送到 #DrillStatus.TaskIO
   IF #EdgeDetc.Pulse[0] AND NOT (#MainStep.S15) THEN
       #DrillStatus.TaskIO := FALSE;
   END_IF;
   // 含义：条件 #EdgeDetc.Pulse[0] AND NOT (#MainStep.S15) 成立时，将 FALSE 传送到 #DrillStatus.TaskNIO
   IF #EdgeDetc.Pulse[0] AND NOT (#MainStep.S15) THEN
       #DrillStatus.TaskNIO := FALSE;
   END_IF;
   // 含义：将 (#EdgeDetc.Pulse[0] AND NOT ("DB1060_AutoStep".HorDrillAutoStep.HorDrillStep.Busy)) OR (#EdgeDetc.Pulse[0] AND #MainStep.S15) 赋给 #MainStep.S15
   #MainStep.S15 := (#EdgeDetc.Pulse[0] AND NOT ("DB1060_AutoStep".HorDrillAutoStep.HorDrillStep.Busy)) OR (#EdgeDetc.Pulse[0] AND #MainStep.S15);

   // ---------- 网络 11 ----------
   // 标题：***************************水平钻孔开始*****************************
   // 含义：条件 #MainStep.S15 AND NOT (#MainStep.S20) 成立时，将 TRUE 传送到 "DB1060_AutoStep".HorDrillAutoStep.HorDrillStep.StartCmd
   IF #MainStep.S15 AND NOT (#MainStep.S20) THEN
       "DB1060_AutoStep".HorDrillAutoStep.HorDrillStep.StartCmd := TRUE;
   END_IF;
   // 含义：条件 ((#MainStep.S15 AND NOT (#MainStep.S20)) AND "DB1060_AutoStep".HorDrillAutoStep.HorDrillStep.TaskDone) AND "DB1060_AutoStep".HorDrillAutoStep.HorDrillStep.TaskIO 成立时，将 TRUE 传送到 #DrillStatus.TaskIO
   IF ((#MainStep.S15 AND NOT (#MainStep.S20)) AND "DB1060_AutoStep".HorDrillAutoStep.HorDrillStep.TaskDone) AND "DB1060_AutoStep".HorDrillAutoStep.HorDrillStep.TaskIO THEN
       #DrillStatus.TaskIO := TRUE;
   END_IF;
   // 含义：条件 ((#MainStep.S15 AND NOT (#MainStep.S20)) AND "DB1060_AutoStep".HorDrillAutoStep.HorDrillStep.TaskDone) AND "DB1060_AutoStep".HorDrillAutoStep.HorDrillStep.TaskNIO 成立时，将 TRUE 传送到 #DrillStatus.TaskNIO
   IF ((#MainStep.S15 AND NOT (#MainStep.S20)) AND "DB1060_AutoStep".HorDrillAutoStep.HorDrillStep.TaskDone) AND "DB1060_AutoStep".HorDrillAutoStep.HorDrillStep.TaskNIO THEN
       #DrillStatus.TaskNIO := TRUE;
   END_IF;
   // 含义：将 (#MainStep.S15 AND "DB1060_AutoStep".HorDrillAutoStep.HorDrillStep.TaskDone) OR (#MainStep.S15 AND #MainStep.S20) 赋给 #MainStep.S20
   #MainStep.S20 := (#MainStep.S15 AND "DB1060_AutoStep".HorDrillAutoStep.HorDrillStep.TaskDone) OR (#MainStep.S15 AND #MainStep.S20);

   // ---------- 网络 12 ----------
   // 标题：钻孔结束
   // 含义：条件 #MainStep.S20 AND NOT (#MainStep.S25) 成立时，将 TRUE 传送到 #DrillStatus.TaskDone
   IF #MainStep.S20 AND NOT (#MainStep.S25) THEN
       #DrillStatus.TaskDone := TRUE;
   END_IF;
   // 含义：将 (#MainStep.S20 AND NOT (#Cmd.Auto.Drill)) OR (#MainStep.S20 AND #MainStep.S25) 赋给 #MainStep.S25
   #MainStep.S25 := (#MainStep.S20 AND NOT (#Cmd.Auto.Drill)) OR (#MainStep.S20 AND #MainStep.S25);

   // ---------- 网络 13 ----------
   // 标题：检查机器人状态
   // 含义：条件 #EdgeDetc.Pulse[0] AND NOT (#MainStep.S40) 成立时，将 TRUE 传送到 #DrillStatus.Busy
   IF #EdgeDetc.Pulse[0] AND NOT (#MainStep.S40) THEN
       #DrillStatus.Busy := TRUE;
   END_IF;
   // 含义：条件 #EdgeDetc.Pulse[0] AND NOT (#MainStep.S40) 成立时，将 FALSE 传送到 #DrillStatus.TaskIO
   IF #EdgeDetc.Pulse[0] AND NOT (#MainStep.S40) THEN
       #DrillStatus.TaskIO := FALSE;
   END_IF;
   // 含义：条件 #EdgeDetc.Pulse[0] AND NOT (#MainStep.S40) 成立时，将 FALSE 传送到 #DrillStatus.TaskNIO
   IF #EdgeDetc.Pulse[0] AND NOT (#MainStep.S40) THEN
       #DrillStatus.TaskNIO := FALSE;
   END_IF;
   // 含义：将 (#EdgeDetc.Pulse[0] AND NOT ("DB1060_AutoStep".DownDrillAutoStep.DownDrillStep.Busy)) OR (#EdgeDetc.Pulse[0] AND #MainStep.S45) 赋给 #MainStep.S45
   #MainStep.S45 := (#EdgeDetc.Pulse[0] AND NOT ("DB1060_AutoStep".DownDrillAutoStep.DownDrillStep.Busy)) OR (#EdgeDetc.Pulse[0] AND #MainStep.S45);

   // ---------- 网络 14 ----------
   // 标题：***************************向下钻孔开始*****************************
   // 含义：条件 #MainStep.S45 AND NOT (#MainStep.S50) 成立时，将 TRUE 传送到 "DB1060_AutoStep".DownDrillAutoStep.DownDrillStep.StartCmd
   IF #MainStep.S45 AND NOT (#MainStep.S50) THEN
       "DB1060_AutoStep".DownDrillAutoStep.DownDrillStep.StartCmd := TRUE;
   END_IF;
   // 含义：条件 ((#MainStep.S45 AND NOT (#MainStep.S50)) AND "DB1060_AutoStep".DownDrillAutoStep.DownDrillStep.TaskDone) AND "DB1060_AutoStep".DownDrillAutoStep.DownDrillStep.TaskIO 成立时，将 TRUE 传送到 #DrillStatus.TaskIO
   IF ((#MainStep.S45 AND NOT (#MainStep.S50)) AND "DB1060_AutoStep".DownDrillAutoStep.DownDrillStep.TaskDone) AND "DB1060_AutoStep".DownDrillAutoStep.DownDrillStep.TaskIO THEN
       #DrillStatus.TaskIO := TRUE;
   END_IF;
   // 含义：条件 ((#MainStep.S45 AND NOT (#MainStep.S50)) AND "DB1060_AutoStep".DownDrillAutoStep.DownDrillStep.TaskDone) AND "DB1060_AutoStep".DownDrillAutoStep.DownDrillStep.TaskNIO 成立时，将 TRUE 传送到 #DrillStatus.TaskNIO
   IF ((#MainStep.S45 AND NOT (#MainStep.S50)) AND "DB1060_AutoStep".DownDrillAutoStep.DownDrillStep.TaskDone) AND "DB1060_AutoStep".DownDrillAutoStep.DownDrillStep.TaskNIO THEN
       #DrillStatus.TaskNIO := TRUE;
   END_IF;
   // 含义：将 (#MainStep.S45 AND "DB1060_AutoStep".DownDrillAutoStep.DownDrillStep.TaskDone) OR (#MainStep.S45 AND #MainStep.S50) 赋给 #MainStep.S50
   #MainStep.S50 := (#MainStep.S45 AND "DB1060_AutoStep".DownDrillAutoStep.DownDrillStep.TaskDone) OR (#MainStep.S45 AND #MainStep.S50);

   // ---------- 网络 15 ----------
   // 标题：钻孔结束
   // 含义：条件 #MainStep.S50 AND NOT (#MainStep.S52) 成立时，将 TRUE 传送到 #DrillStatus.TaskDone
   IF #MainStep.S50 AND NOT (#MainStep.S52) THEN
       #DrillStatus.TaskDone := TRUE;
   END_IF;
   // 含义：将 (#MainStep.S50 AND NOT (#Cmd.Auto.Drill)) OR (#MainStep.S50 AND #MainStep.S52) 赋给 #MainStep.S52
   #MainStep.S52 := (#MainStep.S50 AND NOT (#Cmd.Auto.Drill)) OR (#MainStep.S50 AND #MainStep.S52);

   // ---------- 网络 16 ----------
   // 标题：检查机器人状态
   // 含义：条件 #EdgeDetc.Pulse[0] AND NOT (#MainStep.S55) 成立时，将 TRUE 传送到 #DrillStatus.Busy
   IF #EdgeDetc.Pulse[0] AND NOT (#MainStep.S55) THEN
       #DrillStatus.Busy := TRUE;
   END_IF;
   // 含义：条件 #EdgeDetc.Pulse[0] AND NOT (#MainStep.S55) 成立时，将 FALSE 传送到 #CheckBitStatus.TaskIO
   IF #EdgeDetc.Pulse[0] AND NOT (#MainStep.S55) THEN
       #CheckBitStatus.TaskIO := FALSE;
   END_IF;
   // 含义：条件 #EdgeDetc.Pulse[0] AND NOT (#MainStep.S55) 成立时，将 FALSE 传送到 #CheckBitStatus.TaskNIO
   IF #EdgeDetc.Pulse[0] AND NOT (#MainStep.S55) THEN
       #CheckBitStatus.TaskNIO := FALSE;
   END_IF;
   // 含义：将 (#EdgeDetc.Pulse[0] AND NOT ("DB720_KuKa_MainCtrl".CheckBit.Busy)) OR (#EdgeDetc.Pulse[0] AND #MainStep.S55) 赋给 #MainStep.S55
   #MainStep.S55 := (#EdgeDetc.Pulse[0] AND NOT ("DB720_KuKa_MainCtrl".CheckBit.Busy)) OR (#EdgeDetc.Pulse[0] AND #MainStep.S55);

   // ---------- 网络 17 ----------
   // 标题：****************************校验批头*******************************
   // 含义：条件 #MainStep.S55 AND NOT (#MainStep.S57) 成立时，将 TRUE 传送到 "DB720_KuKa_MainCtrl".CheckBit.StartCmd
   IF #MainStep.S55 AND NOT (#MainStep.S57) THEN
       "DB720_KuKa_MainCtrl".CheckBit.StartCmd := TRUE;
   END_IF;
   // 含义：条件 ((#MainStep.S55 AND NOT (#MainStep.S57)) AND "DB720_KuKa_MainCtrl".CheckBit.TaskDone) AND "DB720_KuKa_MainCtrl".CheckBit.TaskIO 成立时，将 TRUE 传送到 #CheckBitStatus.TaskIO
   IF ((#MainStep.S55 AND NOT (#MainStep.S57)) AND "DB720_KuKa_MainCtrl".CheckBit.TaskDone) AND "DB720_KuKa_MainCtrl".CheckBit.TaskIO THEN
       #CheckBitStatus.TaskIO := TRUE;
   END_IF;
   // 含义：条件 ((#MainStep.S55 AND NOT (#MainStep.S57)) AND "DB720_KuKa_MainCtrl".CheckBit.TaskDone) AND "DB720_KuKa_MainCtrl".CheckBit.TaskNIO 成立时，将 TRUE 传送到 #CheckBitStatus.TaskNIO
   IF ((#MainStep.S55 AND NOT (#MainStep.S57)) AND "DB720_KuKa_MainCtrl".CheckBit.TaskDone) AND "DB720_KuKa_MainCtrl".CheckBit.TaskNIO THEN
       #CheckBitStatus.TaskNIO := TRUE;
   END_IF;
   // 含义：将 (#MainStep.S55 AND "DB720_KuKa_MainCtrl".CheckBit.TaskDone) OR (#MainStep.S55 AND #MainStep.S57) 赋给 #MainStep.S57
   #MainStep.S57 := (#MainStep.S55 AND "DB720_KuKa_MainCtrl".CheckBit.TaskDone) OR (#MainStep.S55 AND #MainStep.S57);

   // ---------- 网络 18 ----------
   // 标题：校验结束
   // 含义：条件 #MainStep.S57 AND NOT (#MainStep.S60) 成立时，将 TRUE 传送到 #CheckBitStatus.TaskDone
   IF #MainStep.S57 AND NOT (#MainStep.S60) THEN
       #CheckBitStatus.TaskDone := TRUE;
   END_IF;
   // 含义：将 (#MainStep.S57 AND NOT (#Cmd.Auto.Drill)) OR (#MainStep.S57 AND #MainStep.S60) 赋给 #MainStep.S60
   #MainStep.S60 := (#MainStep.S57 AND NOT (#Cmd.Auto.Drill)) OR (#MainStep.S57 AND #MainStep.S60);

   // ---------- 网络 19 ----------
   // 标题：自动步结束
   // 含义：将 #MainStep.S11 OR #MainStep.S25 OR #MainStep.S52 OR #MainStep.S60 OR #MainStep.ErrEnd 赋给 #MainStep.End
   #MainStep.End := #MainStep.S11 OR #MainStep.S25 OR #MainStep.S52 OR #MainStep.S60 OR #MainStep.ErrEnd;

   // ---------- 网络 20 ----------
   // 标题：节拍显示
   // 含义：当 #MainStep.S1 为 TRUE 时置位 #CycleTime.StepStart，否则复位（触点→线圈）
   IF #MainStep.S1 THEN
       #CycleTime.StepStart := TRUE;
   ELSE
       #CycleTime.StepStart := FALSE;
   END_IF;
   // 含义：调用块/实例 #CycleTime
   #CycleTime();

   // ---------- 网络 21 ----------
   // 含义：将 0 赋给 #AtCmd
   #AtCmd := 0;

   // ---------- 网络 22 ----------
   // （空白网络）
END_FUNCTION_BLOCK

